// TIA Portal project "261019_Kommissionierung_GA_Analog2_20261019_1400" (V17)

(* hardware
DEVICE "S7300/ET200M-Station_1"  S7-300 station
   slot 0: "Profilschiene_0"  Rail  6ES7 390-1***0-0AA0
   slot 1: "PS 307 5A_1"  PS 307 5A  6ES7 307-1EA01-0AA0
   slot 2: "PLC_WBS_Bus_1"  CPU 314C-2 DP  6ES7 314-6CH04-0AB0  V3.3
      slot 0: "MPI-Schnittstelle_1"  MPI
      slot 1: "DP-Schnittstelle_1"  DP
      slot 2: "DI 24/DO 16_1"  DI24/DO16
      slot 3: "AI 5/AO 2_1"  AI5/AO2
      slot 4: "Zählen_1"  Counter
      slot 5: "Positionieren_1"  Positioning
   slot 4: "DI 64x24VDC sinking/souring_1"  DI64 x 24VDC  6ES7 321-1BP00-0AA0
   slot 5: "DI 64x24VDC sinking/souring_2"  DI64 x 24VDC  6ES7 321-1BP00-0AA0
   slot 6: "DI 64x24VDC sinking/souring_3"  DI64 x 24VDC  6ES7 321-1BP00-0AA0
   slot 7: "DI 64x24VDC sinking/souring_4"  DI64 x 24VDC  6ES7 321-1BP00-0AA0
   slot 8: "DO 64x24VDC/0.3A sourcing_1"  DO64 x 24VDC / 0.3A, P  6ES7 322-1BP00-0AA0
   slot 9: "DO 64x24VDC/0.3A sourcing_2"  DO64 x 24VDC / 0.3A, P  6ES7 322-1BP00-0AA0
   slot 10: "DO 64x24VDC/0.3A sourcing_3"  DO64 x 24VDC / 0.3A, P  6ES7 322-1BP00-0AA0
   slot 11: "DO 64x24VDC/0.3A sourcing_4"  DO64 x 24VDC / 0.3A, P  6ES7 322-1BP00-0AA0
*)

// ===== PLC "PLC_WBS_Bus_1"  CPU 314C-2 DP =====

VAR_GLOBAL   // PLC tag table "Standard-Variablentabelle"
   "NotAusOK" AT %M20.0 : Bool;
   "Band 1 Grün" AT %M41.0 : Bool;
   "Band 2 Blau" AT %M40.1 : Bool;
   "Signal_Start_Bearbeitung" AT %M80.0 : Bool;
   "Band 3 Blau" AT %M40.3 : Bool;
   "Auswahl Unterteil Blau" AT %M42.0 : Bool;
   "Band 6 Blau" AT %M40.4 : Bool;
   "Klemmen UT" AT %M80.2 : Bool;
   "Klemmen Unterteil Blau" AT %M44.0 : Bool;
   "Auswahl Oberteil Blau" AT %M42.1 : Bool;
   "Klemmen Oberteil Blau" AT %M44.1 : Bool;
   "Klemmen OT" AT %M80.3 : Bool;
   "Freigabe_Zusammenbau UT Blau" AT %M82.0 : Bool;
   "Freigabe_Zusammenbau OT Blau" AT %M82.1 : Bool;
   "Teil in Pos. nf" AT %M81.0 : Bool;
   "Teil in Pos. pf" AT %M81.1 : Bool;
   "Z-Achse Greifer Blau" AT %M82.2 : Bool;
   "Greifer Blau" AT %M82.3 : Bool;
   "X-Achse Greifer" AT %M82.4 : Bool;
   "Sensor Weitergabe pf Blau" AT %M82.6 : Bool;
   "Sensor Weitergabe pf 2 Blau" AT %M82.7 : Bool;
   "Start Zusammenbau Blau" AT %M83.0 : Bool;
   "Start zusammen bau pf Blau" AT %M83.3 : Bool;
   "Greifer X-Achse Blau" AT %M83.4 : Bool;
   "Z-Achse senken Zusammenbau" AT %M83.5 : Bool;
   "Teil erkannt pf Blau" AT %M83.7 : Bool;
   "Zusammenbau fertig" AT %M84.6 : Bool;
   "FreigabeKommissionierung Blau" AT %M90.0 : Bool;
   "Anlage Freigegeben" AT %M1.0 : Bool;
   "2Hz" AT %M100.3 : Bool;
   "Betriebsbereit" AT %M20.1 : Bool;
   "Anlage An" AT %M20.2 : Bool;
   "Warnung" AT %M20.3 : Bool;
   "T10s" AT %M20.4 : Bool;
   "Betriebsbereit pf" AT %M20.5 : Bool;
   "Objekt erzeugen Blau" AT %M20.6 : Bool;
   "Start Allgemein" AT %M20.7 : Bool;
   "Start pf" AT %M21.0 : Bool;
   "Auswahl OT_UT Blau" AT %M92.0 : Bool;
   "Start_Signal" AT %M21.2 : Bool;
   "Greifer nf Blau" AT %M83.2 : Bool;
   "X-Achse pf" AT %M84.3 : Bool;
   "Teil erkannt pf(1)" AT %M79.0 : Bool;
   "Start Zusammenbau pf" AT %M81.2 : Bool;
   "Teil fertig Blau" AT %M84.4 : Bool;
   "Grundstellung Roboter Blau" AT %M84.7 : Bool;
   "Teil fertig SR Blau" AT %M85.0 : Bool;
   "Emmit pf" AT %M21.4 : Bool;
   "TB3006 pf" AT %M40.2 : Bool;
   "Start  t1s. pf Blau" AT %M19.1 : Bool;
   "Neues Objekt pf Blau" AT %M19.2 : Bool;
   "Signal_Start_Bearbeitung Grün" AT %M80.1 : Bool;
   "Band 2 Grün" AT %M40.0 : Bool;
   "TB 4006 pf" AT %M40.5 : Bool;
   "Band 3 Grün" AT %M40.6 : Bool;
   "Auswahl Oberteil Grün" AT %M40.7 : Bool;
   "Auswahl Unterteil Grün" AT %M41.1 : Bool;
   "Teil vor Pos. nf" AT %M81.4 : Bool;
   "Klemmen Oberteil Grün" AT %M44.2 : Bool;
   "Teil in Pos. nf Grün" AT %M81.3 : Bool;
   "Klemmen Unterteil Grün" AT %M44.3 : Bool;
   "Band 6 Grün" AT %M41.2 : Bool;
   "FreigabeKommissionierung Grün" AT %M90.1 : Bool;
   "Freigabe_Zusammenbau UT Grün" AT %M84.0 : Bool;
   "Sensor Weitergabe pf Grün" AT %M80.4 : Bool;
   "Freigabe_Zusammenbau OT Grün" AT %M84.1 : Bool;
   "Sensor Weitergabe pf 2 Grün" AT %M84.5 : Bool;
   "Start Zusammenbau Grün" AT %M83.1 : Bool;
   "Start zusammen bau pf Grün" AT %M83.6 : Bool;
   "X-Achse pf Grün" AT %M85.1 : Bool;
   "Z-Achse Greifer Grün" AT %M85.2 : Bool;
   "Greifer X-Achse Grün" AT %M85.3 : Bool;
   "Teil erkannt pf Grün" AT %M85.4 : Bool;
   "Teil erkannt pf(1) Grün" AT %M85.5 : Bool;
   "Teil fertig Grün" AT %M85.6 : Bool;
   "Greifer Grün" AT %M85.7 : Bool;
   "Start Zusammenbau pf Grün" AT %M90.2 : Bool;
   "Greifer nf Grün" AT %M90.3 : Bool;
   "Greifer X-Achse Grün(1)" AT %M90.4 : Bool;
   "Teil erkannt pf Grün(1)" AT %M90.5 : Bool;
   "Teil fertig SR Grün" AT %M90.6 : Bool;
   "Grundstellung Roboter Grün" AT %M90.7 : Bool;
   "FreigabeKommissionierung Grün(1)" AT %M92.1 : Bool;
   "Auswahl OT_UT Grün" AT %M92.2 : Bool;
   "Start  t1s. pf Grün" AT %M19.3 : Bool;
   "Neues Objekt pf Grün" AT %M19.4 : Bool;
   "Objekt erzeugen Grün" AT %M19.5 : Bool;
END_VAR

VAR_GLOBAL   // PLC tag table "Betriebsart"
   "S0_HS" AT %E0.0 : Bool;   // Hauptschalter 0-Aus, 1-Ein
   "S1_Not_Halt" AT %E0.1 : Bool;   // Not-Halt NC
   "S2_START" AT %E0.2 : Bool;   // Taster START NO
   "S3_STOP" AT %E0.3 : Bool;   // Taster STOP NC
   "Res_E04" AT %E0.4 : Bool;
   "Res_E05" AT %E0.5 : Bool;
   "Res_E06" AT %E0.6 : Bool;
   "Res_E07" AT %E0.7 : Bool;
   "Res_E10" AT %E1.0 : Bool;
   "Res_E11" AT %E1.1 : Bool;
   "Res_E12" AT %E1.2 : Bool;
   "Res_E13" AT %E1.3 : Bool;
   "Res_E14" AT %E1.4 : Bool;
   "Res_E15" AT %E1.5 : Bool;
   "Res_E16" AT %E1.6 : Bool;
   "Factory_IO_RUN" AT %E1.7 : Bool;   // Rückmeldung Factory IO läuft
   "P1_MS_RT" AT %A0.0 : Bool;   // Meldesäule Rot
   "P2_MS_GE" AT %A0.1 : Bool;   // Meldesäule Gelb
   "P3_MS_GN" AT %A0.2 : Bool;   // Meldesäule Grün
   "P10_START" AT %A0.3 : Bool;   // Anzeige grün in START-Taster
   "P11_STOP" AT %A0.4 : Bool;   // Anzeige gelb in START-Taster
   "Res_A0.5" AT %A0.5 : Bool;
   "P12_Anfahrwarnung" AT %A0.6 : Bool;   // Rundumleuchte System
   "P13_Sirene" AT %A0.7 : Bool;   // Sirene System
   "Res_A10" AT %A1.0 : Bool;
   "Res_A11" AT %A1.1 : Bool;
   "Res_A12" AT %A1.2 : Bool;
   "Res_A13" AT %A1.3 : Bool;
   "Res_A14" AT %A1.4 : Bool;
   "Res_A15" AT %A1.5 : Bool;
   "Res_A16" AT %A1.6 : Bool;
   "Res_A17" AT %A1.7 : Bool;
   "Log_1" AT %M0.1 : Bool;   // statisch "1"
   "Log_0" AT %M0.0 : Bool;   // statisch "0"
   "Takt_1HZ" AT %M100.5 : Bool;   // Taktmerker 1 Hz
   "Anzeige_Anzahl_Teile_BL" AT %AW22 : Int;   // Anzeige Teile blau im Lager
   "Anzeige_Anzahl_Teile_GN" AT %AW24 : Int;   // Anzeige Teile grün im Lager
   "Reset Nothalt" AT %M0.2 : Bool;
END_VAR

VAR_GLOBAL   // PLC tag table "Montage"
   "B3001_TB3001" AT %E2.0 : Bool;   // Transportband-Ende NC
   "B3002_TB3001" AT %E2.1 : Bool;   // Teil nachPositionierer NC
   "B3003_Teil_vor_POS" AT %E2.2 : Bool;   // Teil vor Positionierer NC
   "B3004_TB3001" AT %E2.3 : Bool;   // Transportband-Anfang NC
   "B3005_TB3002" AT %E2.4 : Bool;   // Transportband-Ende NC
   "B3006_TB3006" AT %E2.5 : Bool;   // Teil vor Schwenkarm NC
   "B3007_UT_BL" AT %E2.6 : Bool;   // Farbsensor Erkennung Farbteil Unterteil blau
   "B3008_OT_BL" AT %E2.7 : Bool;   // Farbsensor Erkennung Farbteil Oberteil blau
   "B3009_TB3006" AT %E3.0 : Bool;   // Transportband-Anfang NC
   "B3010_TB3007" AT %E3.1 : Bool;   // Transportband-Ende NC
   "B3011_TB3007" AT %E3.2 : Bool;   // Transportband-Anfang NC
   "B3012_TB3008" AT %E3.3 : Bool;   // Transportband-Ende NC
   "B3013_TB3008" AT %E3.4 : Bool;   // Transportband-Anfang NC
   "B3014_TB3005" AT %E3.5 : Bool;   // Transportband-Anfang NC
   "B3015_TB3005" AT %E3.6 : Bool;   // Transportband-Ende
   "B3016_TB3004" AT %E3.7 : Bool;   // Transportband-Anfang
   "B3017_Teil_vor_POS" AT %E4.0 : Bool;   // Teil vor Positionierer NC
   "B3018_TB3004" AT %E4.1 : Bool;   // Transportband-Ende NC
   "B3030_POS3001_geklemmt" AT %E4.2 : Bool;   // Positionierer RM geklemmt
   "B3031_POS3001_Heben_Senken" AT %E4.3 : Bool;   // Positionierer RM Bewegung
   "B3040_POS3002_geklemmt" AT %E4.4 : Bool;   // Positionierer RM geklemmt
   "B3041_POS3002_Heben_Senken" AT %E4.5 : Bool;   // Positionierer RM Bewegung
   "Res_E46" AT %E4.6 : Bool;
   "Res_E47" AT %E4.7 : Bool;
   "B3050_PAP3001_RM_X" AT %E5.0 : Bool;
   "B3051_PAP3001_RM_Z" AT %E5.1 : Bool;
   "B3052_PAP3001_Teil_erkannt" AT %E5.2 : Bool;
   "B3070_FZ_3001_Busy" AT %E5.3 : Bool;
   "B3071_FZ_3001_Error" AT %E5.4 : Bool;
   "B3072_FZ_Tür_offen" AT %E5.5 : Bool;
   "Res_E56" AT %E5.6 : Bool;
   "Res_E57" AT %E5.7 : Bool;
   "B4001_TB4001" AT %E6.0 : Bool;   // Transportband-Ende NC
   "B4002_TB4001" AT %E6.1 : Bool;   // Teil nachPositionierer NC
   "B4003_Teil_vor_POS" AT %E6.2 : Bool;   // Teil vor Positionierer NC
   "B4004_TB4001" AT %E6.3 : Bool;   // Transportband-Anfang NC
   "B4005_TB4002" AT %E6.4 : Bool;   // Transportband-Ende NC
   "B4006_TB4006" AT %E6.5 : Bool;   // Teil vor Schwenkarm NC
   "B4007_UT_GN" AT %E6.6 : Bool;   // Farbsensor Erkennung Farbteil Unterteil blau
   "B4008_OT_GN" AT %E6.7 : Bool;   // Farbsensor Erkennung Farbteil Oberteil blau
   "B4009_TB4006" AT %E7.0 : Bool;   // Transportband-Anfang NC
   "B4010_TB4007" AT %E7.1 : Bool;   // Transportband-Ende NC
   "B4011_TB4007" AT %E7.2 : Bool;   // Transportband-Anfang NC
   "B4012_TB4008" AT %E7.3 : Bool;   // Transportband-Ende NC
   "B4013_TB4008" AT %E7.4 : Bool;   // Transportband-Anfang NC
   "B4014_TB4005" AT %E7.5 : Bool;   // Transportband-Anfang NC
   "B4015_TB4005" AT %E7.6 : Bool;   // Transportband-Ende
   "B4016_TB4004" AT %E7.7 : Bool;   // Transportband-Anfang
   "B4017_Teil_vor_POS" AT %E8.0 : Bool;   // Teil vor Positionierer NC
   "B4018_TB4004" AT %E8.1 : Bool;   // Transportband-Ende NC
   "B4030_POS4001_geklemmt" AT %E8.2 : Bool;   // Positionierer RM geklemmt
   "B4031_POS4001_Heben_Senken" AT %E8.3 : Bool;   // Positionierer RM Bewegung
   "B4040_POS4002_geklemmt" AT %E8.4 : Bool;   // Positionierer RM geklemmt
   "B4041_POS4002_Heben_Senken" AT %E8.5 : Bool;   // Positionierer RM Bewegung
   "Res_E86" AT %E8.6 : Bool;
   "Res_E87" AT %E8.7 : Bool;
   "B4050_PAP4001_RM_X" AT %E9.0 : Bool;   // Pick-and-Place X-aktiv
   "B4051_PAP4001_RM_Z" AT %E9.1 : Bool;   // Pick-and-Place Z-aktiv
   "B4052_PAP4001_Teil_erkannt" AT %E9.2 : Bool;   // Teil am Greifer erkannt
   "B4070_FZ_4001_Busy" AT %E9.3 : Bool;   // Fertigungszentrum
   "B4071_FZ_4001_Error" AT %E9.4 : Bool;   // Fertigungszentrum
   "B4072_FZ_4001_Tür_offen" AT %E9.5 : Bool;   // Fertigungszentrum
   "Res_E96" AT %E9.6 : Bool;
   "Res_E97" AT %E9.7 : Bool;
   "TB3001" AT %A2.0 : Bool;
   "TB3002" AT %A2.1 : Bool;
   "TB3003" AT %A2.2 : Bool;
   "TB3004" AT %A2.3 : Bool;
   "TB3005" AT %A2.4 : Bool;
   "TB3006" AT %A2.5 : Bool;
   "TB3007" AT %A2.6 : Bool;
   "TB3008" AT %A2.7 : Bool;
   "FZ_3001_Start" AT %A3.0 : Bool;   // Fertigungszentrum Start
   "FZ_3001_Stop" AT %A3.1 : Bool;   // Fertigungszentrum Stop
   "FZ_3001_OT_UT" AT %A3.2 : Bool;   // Fertigungszentrum UT =0 / OT=1
   "Sorter_Arm_3001_schwenken" AT %A3.3 : Bool;
   "Sorter_Arm_3001_Band_V" AT %A3.4 : Bool;
   "Sorter_Arm_3001_Band_R" AT %A3.5 : Bool;
   "POS3001_Klemmen" AT %A3.6 : Bool;
   "POS3001_Heben" AT %A3.7 : Bool;
   "POS3002_Klemmen" AT %A4.0 : Bool;
   "POS3002_Heben" AT %A4.1 : Bool;
   "PAP3001_X" AT %A4.2 : Bool;
   "PAP3001_Z" AT %A4.3 : Bool;
   "PAP3001_Greifer" AT %A4.4 : Bool;
   "STOP_3001" AT %A4.5 : Bool;
   "Res_A46" AT %A4.6 : Bool;
   "Emitter_1 Blau" AT %A4.7 : Bool;   // Emitter_1
   "TB4001" AT %A5.0 : Bool;
   "TB4002" AT %A5.1 : Bool;
   "TB4003" AT %A5.2 : Bool;
   "TB4004" AT %A5.3 : Bool;
   "TB4005" AT %A5.4 : Bool;
   "TB4006" AT %A5.5 : Bool;
   "TB4007" AT %A5.6 : Bool;
   "TB4008" AT %A5.7 : Bool;
   "FZ_4001_Start" AT %A6.0 : Bool;   // Fertigungszentrum Start
   "FZ_4001_Stop" AT %A6.1 : Bool;   // Fertigungszentrum Stop
   "FZ_4001_OT_UT" AT %A6.2 : Bool;   // Fertigungszentrum UT =0 / OT=1
   "Sorter_Arm_4001_schwenken" AT %A6.3 : Bool;
   "Sorter_Arm_4001_Band_V" AT %A6.4 : Bool;
   "Sorter_Arm_4001_Band_R" AT %A6.5 : Bool;
   "POS4001_Klemmen" AT %A6.6 : Bool;
   "POS4001_Heben" AT %A6.7 : Bool;
   "POS4002_Klemmen" AT %A7.0 : Bool;
   "POS4002_Heben" AT %A7.1 : Bool;
   "PAP4001_X" AT %A7.2 : Bool;
   "PAP4001_Z" AT %A7.3 : Bool;
   "PAP4001_Greifer" AT %A7.4 : Bool;
   "STOP4001" AT %A7.5 : Bool;
   "Res_A76" AT %A7.6 : Bool;
   "Emitter_2 Grün" AT %A7.7 : Bool;
   "FZ_3001_Bearbeitungszeit" AT %EW20 : Int;
   "FZ_4001_Bearbeitungszeit" AT %EW22 : Int;
END_VAR

VAR_GLOBAL   // PLC tag table "Kommisionierung"
   "B5001_TB5001" AT %E10.0 : Bool;   // Teil vom Emitter vorhanden
   "B5002_TB5001" AT %E10.1 : Bool;   // Transportband-Ende
   "B5003_TB5002" AT %E10.2 : Bool;   // Transportband-Anfang
   "B5004_TB5002" AT %E10.3 : Bool;   // Transportband-Ende
   "B5005_TB5003" AT %E10.4 : Bool;   // Transportband-Anfang
   "B5006_TB5003" AT %E10.5 : Bool;   // Transportband-Ende
   "B5007_TB5004" AT %E10.6 : Bool;   // Transportband-Anfang
   "B5008_TB5004" AT %E10.7 : Bool;   // Transportband-Ende
   "B5009_TB5005" AT %E11.0 : Bool;   // Transportband-Anfang
   "B5010_TB5005" AT %E11.1 : Bool;   // Transportband-Ende
   "B5011_Farbteil_GN" AT %E11.2 : Bool;   // Farberkennung GN
   "B5012_Farbteil_BL" AT %E11.3 : Bool;   // Farberkennung_BL
   "B5013_TB5006" AT %E11.4 : Bool;   // Transportband-Anfang
   "B5014_TB5006" AT %E11.5 : Bool;   // Transportband-Ende blaue Produkte
   "B5016_Teil_vorhanden" AT %E11.7 : Bool;   // Teil vom Emitter generiert
   "B5018_Teil_vorhanden" AT %E12.1 : Bool;   // Teil vom Emitter generiert
   "B5019_TB5009" AT %E12.2 : Bool;   // Transportband-Anfang
   "B5020_TB5009" AT %E12.3 : Bool;   // Transportband-Ende
   "B5021_TB5010" AT %E12.4 : Bool;   // Transportband-Anfang
   "B5022_TB5010" AT %E12.5 : Bool;   // Transportband-Ende grüne Produkte
   "Res_E126" AT %E12.6 : Bool;
   "Res_E127" AT %E12.7 : Bool;
   "B5030_PAP5001_RM_X" AT %E13.0 : Bool;
   "B5031_PAP5001_RM_Z" AT %E13.1 : Bool;
   "B5032_PAP5001_Teil_erkannt" AT %E13.2 : Bool;
   "B5040_PAP5002_RM_X" AT %E13.3 : Bool;
   "B5041_PAP5002_RM_Z" AT %E13.4 : Bool;
   "B5042_PAP5002_Teil_erkannt" AT %E13.5 : Bool;
   "Res_E136" AT %E13.6 : Bool;
   "Res_E137" AT %E13.7 : Bool;
   "TB5001" AT %A8.0 : Bool;
   "TB5002" AT %A8.1 : Bool;
   "TB5003" AT %A8.2 : Bool;
   "TB5004" AT %A8.3 : Bool;
   "TB5005" AT %A8.4 : Bool;
   "TB5006" AT %A8.5 : Bool;
   "TB5007" AT %A8.6 : Bool;
   "TB5008" AT %A8.7 : Bool;
   "TB5009" AT %A9.0 : Bool;
   "TB5010" AT %A9.1 : Bool;
   "STOP5001" AT %A9.2 : Bool;   // Stopper
   "STOP5002" AT %A9.3 : Bool;   // Stopper
   "STOP5003" AT %A9.4 : Bool;   // Stopper
   "STOP5004" AT %A9.5 : Bool;   // Stopper
   "STOP5005" AT %A9.6 : Bool;   // Stopper
   "Res_A97" AT %A9.7 : Bool;
   "PAP5001_X" AT %A10.0 : Bool;
   "PAP5001_Z" AT %A10.1 : Bool;
   "PAP5001_Greifer" AT %A10.2 : Bool;
   "PAP5002_X" AT %A10.3 : Bool;
   "PAP5002_Z" AT %A10.4 : Bool;
   "PAP5002_Greifer" AT %A10.5 : Bool;
   "Res_A106" AT %A10.6 : Bool;
   "Res_A107" AT %A10.7 : Bool;
   "RS5001_V" AT %A11.0 : Bool;   // Rollensorter Antrieb ein
   "RS5001_links" AT %A11.1 : Bool;   // Rollensorter Steuerung links
   "RS5001_rechts" AT %A11.2 : Bool;   // Rollensorter Steuerung rechts
   "Res_A113" AT %A11.3 : Bool;
   "Res_A114" AT %A11.4 : Bool;
   "Emitter_1" AT %A11.5 : Bool;
   "Emitter_2" AT %A11.6 : Bool;
   "Emitter_3" AT %A11.7 : Bool;
   "TA_P&P2_SetPoint_X" AT %AW24 : Int;
   "TA_P&P2_SetPoint_Z" AT %AW26 : Int;
   "TA_P&P1_SetPoint_X" AT %AW20 : Int;
   "TA_P&P1_SetPoint_Z" AT %AW22 : Int;
   "TA_P&P2_Pos_X" AT %EW24 : Int;
   "TA_P&P2_Pos_Z" AT %EW26 : Int;
   "TA_P&P1_Pos_X" AT %EW20 : Int;
   "TA_P&P1_Pos_Z" AT %EW22 : Int;
   "B5015_Teil_in_Pos" AT %E11.6 : Bool;
   "B5017_Teil_in_Pos" AT %E12.0 : Bool;
END_VAR

// folder: Kommissionierung

DATA_BLOCK "100_DB_Kommissionierung"   // DB100
{ S7_Optimized_Access := 'FALSE' }
VERSION : 0.1
   VAR
      xNotAusOK : Bool;
      xAnlageAusgeschaltet : Bool;
      xAnlageStartet : Bool;
      xAnlageEin : Bool;
      xGA1_Fertig : Bool;
      xGA2_Fertig : Bool;
      strGA1_Meldung : String[30];
      strGA2_Meldung : String[30];
      iIndex_Förderband : Int;
   END_VAR
BEGIN
END_DATA_BLOCK

// folder: Kommissionierung/iDB

DATA_BLOCK "02_AnlageEinAus_DB"   // DB29
{ S7_Optimized_Access := 'FALSE' }
VERSION : 0.1
// stored: InstanceOfName 02_AnlageEinAus
"02_AnlageEinAus"
BEGIN
END_DATA_BLOCK

DATA_BLOCK "03_Förderband_DB"   // DB30
{ S7_Optimized_Access := 'FALSE' }
VERSION : 0.1
// stored: InstanceOfName 03_Förderband
"03_Förderband"
BEGIN
END_DATA_BLOCK

DATA_BLOCK "04_Greifarm_DB"   // DB31
{ S7_Optimized_Access := 'FALSE' }
VERSION : 0.1
// stored: InstanceOfName 04_Greifarm
"04_Greifarm"
BEGIN
END_DATA_BLOCK

DATA_BLOCK "04_Greifarm_DB_1"   // DB32
{ S7_Optimized_Access := 'FALSE' }
VERSION : 0.1
// stored: InstanceOfName 04_Greifarm
"04_Greifarm"
BEGIN
END_DATA_BLOCK

// folder: Montage/Bearbeitung Blau

DATA_BLOCK "01_Transportband vor Bearbeitung_DB"   // DB1
{ S7_Optimized_Access := 'FALSE' }
VERSION : 0.1
// stored: InstanceOfName 01Transportband vor Bearbeitung
"01Transportband vor Bearbeitung"
BEGIN
END_DATA_BLOCK

DATA_BLOCK "Bearbeitung_DB"   // DB2
{ S7_Optimized_Access := 'FALSE' }
VERSION : 0.1
// stored: InstanceOfName 02_Bearbeitung
"02_Bearbeitung"
BEGIN
END_DATA_BLOCK

DATA_BLOCK "02_Bearbeitung_DB"   // DB3
{ S7_Optimized_Access := 'FALSE' }
VERSION : 0.1
// stored: InstanceOfName 02_Bearbeitung
"02_Bearbeitung"
BEGIN
END_DATA_BLOCK

DATA_BLOCK "03_Weiterverarbeitung_DB"   // DB4
{ S7_Optimized_Access := 'FALSE' }
VERSION : 0.1
// stored: InstanceOfName 03_Weiterverarbeitung
"03_Weiterverarbeitung"
BEGIN
END_DATA_BLOCK

DATA_BLOCK "04_Zusammenbau_DB"   // DB6
{ S7_Optimized_Access := 'FALSE' }
VERSION : 0.1
// stored: InstanceOfName 04_Zusammenbau
"04_Zusammenbau"
BEGIN
END_DATA_BLOCK

DATA_BLOCK "05_Weitergabe_DB"   // DB11
{ S7_Optimized_Access := 'FALSE' }
VERSION : 0.1
// stored: InstanceOfName 05_Weitergabe
"05_Weitergabe"
BEGIN
END_DATA_BLOCK

DATA_BLOCK "06_Auswahl OT_UT_DB"   // DB15
{ S7_Optimized_Access := 'FALSE' }
VERSION : 0.1
// stored: InstanceOfName 06_Auswahl OT_UT
"06_Auswahl OT_UT"
BEGIN
END_DATA_BLOCK

// folder: Montage/Bearbeitung Grün

DATA_BLOCK "01_Transportband vor Bearbeitung_DB_Grün"   // DB20
{ S7_Optimized_Access := 'FALSE' }
VERSION : 0.1
// stored: InstanceOfName 01Transportband vor Bearbeitung Grün
"01Transportband vor Bearbeitung Grün"
BEGIN
END_DATA_BLOCK

DATA_BLOCK "Bearbeitung_DB_Grün"   // DB21
{ S7_Optimized_Access := 'FALSE' }
VERSION : 0.1
// stored: InstanceOfName 02_Bearbeitung Grün
"02_Bearbeitung Grün"
BEGIN
END_DATA_BLOCK

DATA_BLOCK "02_Bearbeitung_DB_Grün"   // DB22
{ S7_Optimized_Access := 'FALSE' }
VERSION : 0.1
// stored: InstanceOfName 02_Bearbeitung Grün
"02_Bearbeitung Grün"
BEGIN
END_DATA_BLOCK

DATA_BLOCK "03_Weiterverarbeitung_DB_Grün"   // DB23
{ S7_Optimized_Access := 'FALSE' }
VERSION : 0.1
// stored: InstanceOfName 03_Weiterverarbeitung Grün
"03_Weiterverarbeitung Grün"
BEGIN
END_DATA_BLOCK

DATA_BLOCK "04_Zusammenbau_DB_Grün"   // DB24
{ S7_Optimized_Access := 'FALSE' }
VERSION : 0.1
// stored: InstanceOfName 04_Zusammenbau Grün
"04_Zusammenbau Grün"
BEGIN
END_DATA_BLOCK

DATA_BLOCK "05_Weitergabe_DB_Grün"   // DB25
{ S7_Optimized_Access := 'FALSE' }
VERSION : 0.1
// stored: InstanceOfName 05_Weitergabe Grün
"05_Weitergabe Grün"
BEGIN
END_DATA_BLOCK

DATA_BLOCK "06_Auswahl OT_UT_DB_Grün"   // DB26
{ S7_Optimized_Access := 'FALSE' }
VERSION : 0.1
// stored: InstanceOfName 06_Auswahl OT_UT_Grün
"06_Auswahl OT_UT_Grün"
BEGIN
END_DATA_BLOCK

// folder: Montage/iDB

DATA_BLOCK "05_Weitergabe_DB_1"   // DB5
{ S7_Optimized_Access := 'FALSE' }
VERSION : 0.1
// stored: InstanceOfName 05_Weitergabe
"05_Weitergabe"
BEGIN
END_DATA_BLOCK

DATA_BLOCK "01Transportband vor Bearbeitung Grün_DB"   // DB9
{ S7_Optimized_Access := 'FALSE' }
VERSION : 0.1
// stored: InstanceOfName 01Transportband vor Bearbeitung Grün
"01Transportband vor Bearbeitung Grün"
BEGIN
END_DATA_BLOCK

DATA_BLOCK "02_Bearbeitung Grün_DB"   // DB10
{ S7_Optimized_Access := 'FALSE' }
VERSION : 0.1
// stored: InstanceOfName 02_Bearbeitung Grün
"02_Bearbeitung Grün"
BEGIN
END_DATA_BLOCK

DATA_BLOCK "03_Weiterverarbeitung Grün_DB"   // DB14
{ S7_Optimized_Access := 'FALSE' }
VERSION : 0.1
// stored: InstanceOfName 03_Weiterverarbeitung Grün
"03_Weiterverarbeitung Grün"
BEGIN
END_DATA_BLOCK

DATA_BLOCK "04_Zusammenbau Grün_DB"   // DB16
{ S7_Optimized_Access := 'FALSE' }
VERSION : 0.1
// stored: InstanceOfName 04_Zusammenbau Grün
"04_Zusammenbau Grün"
BEGIN
END_DATA_BLOCK

DATA_BLOCK "05_Weitergabe Grün_DB"   // DB17
{ S7_Optimized_Access := 'FALSE' }
VERSION : 0.1
// stored: InstanceOfName 05_Weitergabe Grün
"05_Weitergabe Grün"
BEGIN
END_DATA_BLOCK

DATA_BLOCK "06_Auswahl OT_UT_Grün_DB"   // DB18
{ S7_Optimized_Access := 'FALSE' }
VERSION : 0.1
// stored: InstanceOfName 06_Auswahl OT_UT_Grün
"06_Auswahl OT_UT_Grün"
BEGIN
END_DATA_BLOCK

DATA_BLOCK "00_Startbedingungen_2_DB"   // DB27
{ S7_Optimized_Access := 'FALSE' }
VERSION : 0.1
// stored: InstanceOfName 00_Startbedingungen_2
"00_Startbedingungen_2"
BEGIN
END_DATA_BLOCK

// folder: (top level)

ORGANIZATION_BLOCK "Main"   // OB1, FBD
TITLE = "Main Program Sweep (Cycle)"
{ S7_Optimized_Access := 'FALSE' }
VERSION : 0.1
   VAR_TEMP
      OB1_EV_CLASS : Byte;   // Bits 0-3 = 1 (Coming event), Bits 4-7 = 1 (Event class 1)
      OB1_SCAN_1 : Byte;   // 1 (Cold restart scan 1 of OB 1), 3 (Scan 2-n of OB 1)
      OB1_PRIORITY : Byte;   // Priority of OB Execution
      OB1_OB_NUMBR : Byte;   // 1 (Organization block 1, OB1)
      OB1_RESERVED_1 : Byte;   // Reserved for system
      OB1_RESERVED_2 : Byte;   // Reserved for system
      OB1_PREV_CYCLE : Int;   // Cycle time of previous OB1 scan (milliseconds)
      OB1_MIN_CYCLE : Int;   // Minimum cycle time of OB1 (milliseconds)
      OB1_MAX_CYCLE : Int;   // Maximum cycle time of OB1 (milliseconds)
      OB1_DATE_TIME : Date_And_Time;   // Date and time OB1 started
   END_VAR
BEGIN

REGION Network 1: Startbedingung
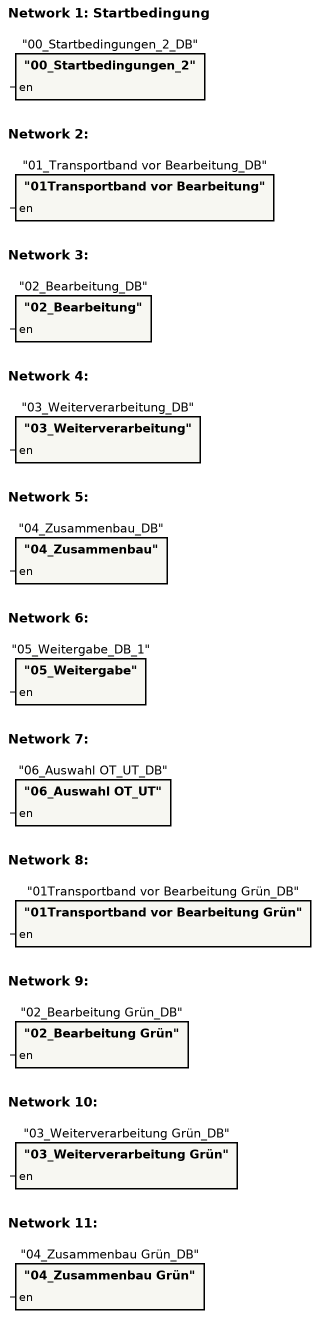
   "00_Startbedingungen_2_DB"();   // "00_Startbedingungen_2"
END_REGION

REGION Network 2
   "01_Transportband vor Bearbeitung_DB"();   // "01Transportband vor Bearbeitung"
END_REGION

REGION Network 3
   "02_Bearbeitung_DB"();   // "02_Bearbeitung"
END_REGION

REGION Network 4
   "03_Weiterverarbeitung_DB"();   // "03_Weiterverarbeitung"
END_REGION

REGION Network 5
   "04_Zusammenbau_DB"();   // "04_Zusammenbau"
END_REGION

REGION Network 6
   "05_Weitergabe_DB_1"();   // "05_Weitergabe"
END_REGION

REGION Network 7
   "06_Auswahl OT_UT_DB"();   // "06_Auswahl OT_UT"
END_REGION

REGION Network 8
   "01Transportband vor Bearbeitung Grün_DB"();   // "01Transportband vor Bearbeitung Grün"
END_REGION

REGION Network 9
   "02_Bearbeitung Grün_DB"();   // "02_Bearbeitung Grün"
END_REGION

REGION Network 10
   "03_Weiterverarbeitung Grün_DB"();   // "03_Weiterverarbeitung Grün"
END_REGION

REGION Network 11
   "04_Zusammenbau Grün_DB"();   // "04_Zusammenbau Grün"
END_REGION

REGION Network 12
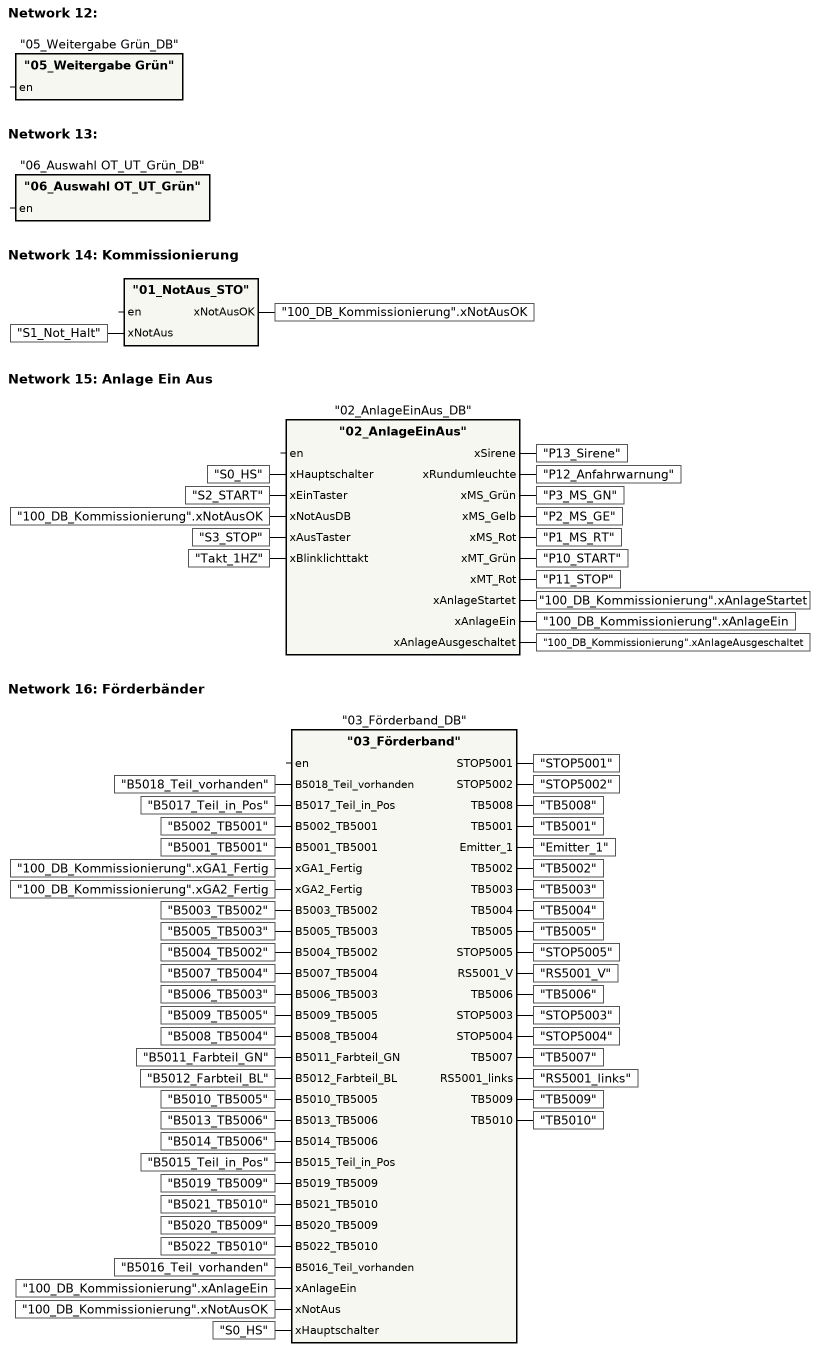
   "05_Weitergabe Grün_DB"();   // "05_Weitergabe Grün"
END_REGION

REGION Network 13
   "06_Auswahl OT_UT_Grün_DB"();   // "06_Auswahl OT_UT_Grün"
END_REGION

REGION Network 14: Kommissionierung
   "01_NotAus_STO"(xNotAus := "S1_Not_Halt", xNotAusOK => "100_DB_Kommissionierung".xNotAusOK);
END_REGION

REGION Network 15: Anlage Ein Aus
   "02_AnlageEinAus_DB"(xHauptschalter := "S0_HS",   // "02_AnlageEinAus"
                        xEinTaster := "S2_START",
                        xNotAusDB := "100_DB_Kommissionierung".xNotAusOK,
                        xAusTaster := "S3_STOP",
                        xBlinklichttakt := "Takt_1HZ",
                        xSirene => "P13_Sirene",
                        xRundumleuchte => "P12_Anfahrwarnung",
                        xMS_Grün => "P3_MS_GN",
                        xMS_Gelb => "P2_MS_GE",
                        xMS_Rot => "P1_MS_RT",
                        xMT_Grün => "P10_START",
                        xMT_Rot => "P11_STOP",
                        xAnlageStartet => "100_DB_Kommissionierung".xAnlageStartet,
                        xAnlageEin => "100_DB_Kommissionierung".xAnlageEin,
                        xAnlageAusgeschaltet => "100_DB_Kommissionierung".xAnlageAusgeschaltet);
END_REGION

REGION Network 16: Förderbänder
   "03_Förderband_DB"(B5018_Teil_vorhanden := "B5018_Teil_vorhanden",   // "03_Förderband"
                      B5017_Teil_in_Pos := "B5017_Teil_in_Pos",
                      B5002_TB5001 := "B5002_TB5001",
                      B5001_TB5001 := "B5001_TB5001",
                      xGA1_Fertig := "100_DB_Kommissionierung".xGA1_Fertig,
                      xGA2_Fertig := "100_DB_Kommissionierung".xGA2_Fertig,
                      B5003_TB5002 := "B5003_TB5002",
                      B5005_TB5003 := "B5005_TB5003",
                      B5004_TB5002 := "B5004_TB5002",
                      B5007_TB5004 := "B5007_TB5004",
                      B5006_TB5003 := "B5006_TB5003",
                      B5009_TB5005 := "B5009_TB5005",
                      B5008_TB5004 := "B5008_TB5004",
                      B5011_Farbteil_GN := "B5011_Farbteil_GN",
                      B5012_Farbteil_BL := "B5012_Farbteil_BL",
                      B5010_TB5005 := "B5010_TB5005",
                      B5013_TB5006 := "B5013_TB5006",
                      B5014_TB5006 := "B5014_TB5006",
                      B5015_Teil_in_Pos := "B5015_Teil_in_Pos",
                      B5019_TB5009 := "B5019_TB5009",
                      B5021_TB5010 := "B5021_TB5010",
                      B5020_TB5009 := "B5020_TB5009",
                      B5022_TB5010 := "B5022_TB5010",
                      B5016_Teil_vorhanden := "B5016_Teil_vorhanden",
                      xAnlageEin := "100_DB_Kommissionierung".xAnlageEin,
                      xNotAus := "100_DB_Kommissionierung".xNotAusOK,
                      xHauptschalter := "S0_HS",
                      STOP5001 => "STOP5001",
                      STOP5002 => "STOP5002",
                      TB5008 => "TB5008",
                      TB5001 => "TB5001",
                      Emitter_1 => "Emitter_1",
                      TB5002 => "TB5002",
                      TB5003 => "TB5003",
                      TB5004 => "TB5004",
                      TB5005 => "TB5005",
                      STOP5005 => "STOP5005",
                      RS5001_V => "RS5001_V",
                      TB5006 => "TB5006",
                      STOP5003 => "STOP5003",
                      STOP5004 => "STOP5004",
                      TB5007 => "TB5007",
                      RS5001_links => "RS5001_links",
                      TB5009 => "TB5009",
                      TB5010 => "TB5010");
END_REGION

REGION Network 17: Greifarm 4
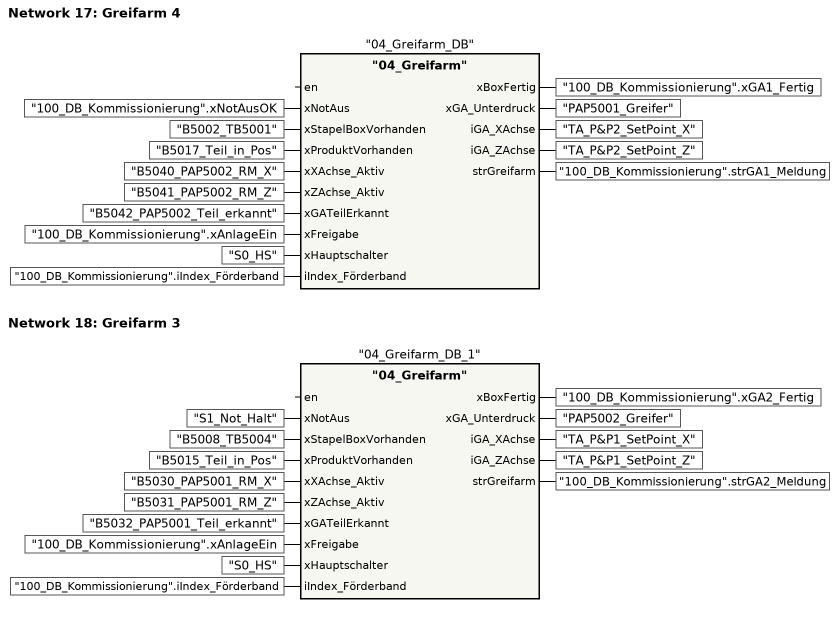
   "04_Greifarm_DB"(xNotAus := "100_DB_Kommissionierung".xNotAusOK,   // "04_Greifarm"
                    xStapelBoxVorhanden := "B5002_TB5001",
                    xProduktVorhanden := "B5017_Teil_in_Pos",
                    xXAchse_Aktiv := "B5040_PAP5002_RM_X",
                    xZAchse_Aktiv := "B5041_PAP5002_RM_Z",
                    xGATeilErkannt := "B5042_PAP5002_Teil_erkannt",
                    xFreigabe := "100_DB_Kommissionierung".xAnlageEin,
                    xHauptschalter := "S0_HS",
                    iIndex_Förderband := "100_DB_Kommissionierung".iIndex_Förderband,
                    xBoxFertig => "100_DB_Kommissionierung".xGA1_Fertig,
                    xGA_Unterdruck => "PAP5001_Greifer",
                    iGA_XAchse => "TA_P&P2_SetPoint_X",
                    iGA_ZAchse => "TA_P&P2_SetPoint_Z",
                    strGreifarm => "100_DB_Kommissionierung".strGA1_Meldung);
END_REGION

REGION Network 18: Greifarm 3
   "04_Greifarm_DB_1"(xNotAus := "S1_Not_Halt",   // "04_Greifarm"
                      xStapelBoxVorhanden := "B5008_TB5004",
                      xProduktVorhanden := "B5015_Teil_in_Pos",
                      xXAchse_Aktiv := "B5030_PAP5001_RM_X",
                      xZAchse_Aktiv := "B5031_PAP5001_RM_Z",
                      xGATeilErkannt := "B5032_PAP5001_Teil_erkannt",
                      xFreigabe := "100_DB_Kommissionierung".xAnlageEin,
                      xHauptschalter := "S0_HS",
                      iIndex_Förderband := "100_DB_Kommissionierung".iIndex_Förderband,
                      xBoxFertig => "100_DB_Kommissionierung".xGA2_Fertig,
                      xGA_Unterdruck => "PAP5002_Greifer",
                      iGA_XAchse => "TA_P&P1_SetPoint_X",
                      iGA_ZAchse => "TA_P&P1_SetPoint_Z",
                      strGreifarm => "100_DB_Kommissionierung".strGA2_Meldung);
END_REGION
END_ORGANIZATION_BLOCK

// folder: Kommissionierung

FUNCTION_BLOCK "03_Förderband"   // FB2, SCL
{ S7_Optimized_Access := 'FALSE' }
VERSION : 0.1
   VAR_INPUT
      B5018_Teil_vorhanden : Bool;
      B5017_Teil_in_Pos : Bool;
      B5002_TB5001 : Bool;
      B5001_TB5001 : Bool;
      xGA1_Fertig : Bool;
      xGA2_Fertig : Bool;
      B5003_TB5002 : Bool;
      B5005_TB5003 : Bool;
      B5004_TB5002 : Bool;
      B5007_TB5004 : Bool;
      B5006_TB5003 : Bool;
      B5009_TB5005 : Bool;
      B5008_TB5004 : Bool;
      B5011_Farbteil_GN : Bool;
      B5012_Farbteil_BL : Bool;
      B5010_TB5005 : Bool;
      B5013_TB5006 : Bool;
      B5014_TB5006 : Bool;
      B5015_Teil_in_Pos : Bool;
      B5019_TB5009 : Bool;
      B5021_TB5010 : Bool;
      B5020_TB5009 : Bool;
      B5022_TB5010 : Bool;
      B5016_Teil_vorhanden : Bool;
      xAnlageEin : Bool;
      xNotAus : Bool;
      xHauptschalter : Bool;
   END_VAR
   VAR_OUTPUT
      STOP5001 : Bool;
      STOP5002 : Bool;
      TB5008 : Bool;
      TB5001 : Bool;
      Emitter_1 : Bool;
      TB5002 : Bool;
      TB5003 : Bool;
      TB5004 : Bool;
      TB5005 : Bool;
      STOP5005 : Bool;
      RS5001_V : Bool;
      TB5006 : Bool;
      STOP5003 : Bool;
      STOP5004 : Bool;
      TB5007 : Bool;
      RS5001_links : Bool;
      TB5009 : Bool;
      TB5010 : Bool;
   END_VAR
   VAR
      stat_iIndex : Int;
      IEC_Timer_0_blau : TON;
      stat_strFörderband : String[15];
      stat_Ntrig1 : Bool;
      stat_Ntig1M : Bool;
      stat_Ntrig2 : Bool;
      stat_Ntig2M : Bool;
      IEC_Timer_1_grün : TON;
   END_VAR
BEGIN
   // ==============================Förderband=======================================
   // Es können zwei verschiedene Produkte über diese Anlage verteilt werden.
   // Blaue oder grüne Produkte.
   // Es darf sich immer nur ein Produkt in der Anlage befinden.

   // Abfrage Hauptschalter
   REGION Abfrage Hauptschalter
       IF NOT #xHauptschalter THEN
           #STOP5001 := 0;
           #STOP5002 := 0;
           #STOP5003 := 0;
           #STOP5004 := 0;
           #STOP5005 := 0;
           #TB5001 := 0;
           #TB5002 := 0;
           #TB5003 := 0;
           #TB5004 := 0;
           #TB5005 := 0;
           #TB5006 := 0;
           #TB5007 := 0;
           #TB5008 := 0;
           #TB5009 := 0;
           #TB5010 := 0;
           #Emitter_1 := 0;
           #RS5001_V := 0;
           #RS5001_links := 0;
           #stat_iIndex := 0;
           #stat_strFörderband := 'HS aus';
           RETURN;
       END_IF;
   END_REGION

   // Abfrage NotAus
   REGION Abfrage NOTAUS
       IF NOT #xNotAus OR "100_DB_Kommissionierung".xAnlageAusgeschaltet THEN
           #STOP5001 := 0;
           #STOP5002 := 0;
           #STOP5003 := 0;
           #STOP5004 := 0;
           #STOP5005 := 0;
           #TB5001 := 0;
           #TB5002 := 0;
           #TB5003 := 0;
           #TB5004 := 0;
           #TB5005 := 0;
           #TB5006 := 0;
           #TB5007 := 0;
           #TB5008 := 0;
           #TB5009 := 0;
           #TB5010 := 0;
           #Emitter_1 := 0;
           #RS5001_V := 0;
           #RS5001_links := 0;
           #stat_iIndex := 0;
           RETURN;
       END_IF;
   END_REGION

   // Entscheidung welches Produkt am Eingang liegt 
   REGION Entscheidung welche Produkt am Eingang liegt
       IF #stat_iIndex = 0 THEN
           #stat_strFörderband := 'Betriebsbereit';
       END_IF;



       IF NOT #B5018_Teil_vorhanden AND #stat_iIndex = 0 AND #xAnlageEin THEN
           #Emitter_1 := 1;
           #STOP5001 := 1;
           #STOP5003 := 1;
           #stat_iIndex := 100;

       END_IF;

       IF NOT #B5016_Teil_vorhanden AND #stat_iIndex = 0 AND #xAnlageEin THEN
           #Emitter_1 := 1;
           #STOP5001 := 1;
           #STOP5003 := 1;
           #stat_iIndex := 200;

       END_IF;
   END_REGION

   // Förderband
   CASE #stat_iIndex OF
       100:    // Stopper ausfahren und Stapelkiste erzeugen
           REGION Stopper ausfahren und Stapelkiste erzeugen

               #STOP5002 := 1;
               #stat_strFörderband := 'In Betrieb';

               // Schritt erhöhen
               IF #B5001_TB5001 THEN
                   #stat_iIndex := #stat_iIndex + 1;
               END_IF;

           END_REGION

       101:    //Förderbänder starten
           REGION Förderbänder starten
               #TB5008 := 1;
               #TB5001 := 1;
               #Emitter_1 := 0;

               IF NOT #B5017_Teil_in_Pos THEN
                   #TB5008 := 0;
               END_IF;


               IF #B5002_TB5001 THEN
                   #TB5001 := 0;
               END_IF; 

               // Zurücksetzen aus vorherigen Schritten
               #Emitter_1 := 0;

               // Schritt erhöhen
               IF NOT #B5017_Teil_in_Pos AND #B5002_TB5001 THEN
                   #stat_iIndex := #stat_iIndex + 1;
               END_IF;
           END_REGION

       102:    // Greifarm abwarten und abtransport über das nächse Förderband
           REGION Greifarm abwarten und abtransport über das nächse Förderband
               IF #xGA1_Fertig THEN
                   (* #STOP5001 := 0; *) // Kann oben bleiben
                   #STOP5002 := 0;
               END_IF;

               IF (* #STOP5001 = 0 AND *) #STOP5002 = 0 THEN
                   #TB5001 := 1;
                   #TB5002 := 1;
               END_IF;

               IF #B5003_TB5002 AND NOT #B5002_TB5001 THEN
                   #TB5001 := 0;
                   #TB5003 := 1;
               END_IF;

               // Schritt erhöhung
               IF NOT #TB5001 AND #TB5002 THEN
                   #stat_iIndex := #stat_iIndex + 1;
               END_IF;
           END_REGION

       103:    // Förderbänder bis zur Farberkennung
           REGION Förderbänder bis zur Farberkennung
               // TB 5002 aus und TB 5003 ein

               IF #B5005_TB5003 AND NOT #B5004_TB5002 THEN
                   #TB5002 := 0;
               END_IF;

               // TB 5003 aus und TB5004 ein
               IF #B5007_TB5004 AND NOT #B5006_TB5003 THEN
                   #TB5003 := 0;
               END_IF;

               IF #B5006_TB5003 THEN
                   #TB5004 := 1;
               END_IF;

               // TB 5004 aus und TB 5005 ein
               IF #B5009_TB5005 AND NOT #B5008_TB5004 THEN
                   #TB5004 := 0;
               END_IF;

               IF #B5008_TB5004 THEN
                   #TB5005 := 1;
               END_IF;

               // Schitt erhöhung
               IF #B5009_TB5005 AND NOT #B5008_TB5004 THEN
                   #stat_iIndex := #stat_iIndex + 1;
               END_IF;

           END_REGION

       104:    // Farberkennung 
           REGION Farberkennung
               // Für blaue Produkte springen wir in 110 
               // Für grüne Produkte springen wir in 210
               IF #B5012_Farbteil_BL THEN
                   #stat_iIndex := 110;
               END_IF;

               IF #B5011_Farbteil_GN THEN
                   #stat_iIndex := 210;
               END_IF;
           END_REGION

       110:    // Rollenförderband blau
           REGION Rollenförderband blau
               #STOP5005 := 1;
               #RS5001_links := 0;
               #RS5001_V := 1;
               #TB5006 := 1;

               IF #B5013_TB5006 AND NOT #B5010_TB5005 THEN
                   #TB5005 := 0;
               END_IF;

               // Flankenauswertung Sensor B5013_TB5006
               // NTrig
               #stat_Ntrig1 := NOT #B5013_TB5006 AND #stat_Ntig1M;
               #stat_Ntig1M := #B5013_TB5006;

               IF #TB5006 = 1 AND #stat_Ntrig1 THEN
                   #STOP5005 := 0;
                   #RS5001_V := 0;
                   #stat_iIndex := #stat_iIndex + 1;
               END_IF;


           END_REGION

       111:    // Remove blaues Produkt 
           REGION Remove blaues Produkt
               #IEC_Timer_0_blau(IN := #B5014_TB5006,
                                     PT := t#0.5s);
                   IF #B5014_TB5006 (* AND #IEC_Timer_0_blau.Q *) THEN
                   #TB5006 := 0;
                   IF NOT #B5015_Teil_in_Pos AND #xAnlageEin THEN
                       #stat_iIndex := 200;
                       #Emitter_1 := 1;
                   ELSE
                       #stat_iIndex := 0;
                   END_IF;
               END_IF;

           END_REGION

       200:    // Stopper ausfahren und Stapelkiste erzeugen
           REGION Stopper ausfahren und Stapelkiste erzeugen

               #STOP5004 := 1;
               #stat_strFörderband := 'In Betrieb';

               // Schritt erhöhen
               IF #B5001_TB5001 THEN
                   #stat_iIndex := #stat_iIndex + 1;
               END_IF;
           END_REGION

       201:    // Förderbänder starten
           REGION Förderbänder starten
               #TB5007 := 1;
               #Emitter_1 := 0;

               IF NOT #B5015_Teil_in_Pos THEN
                   #TB5007 := 0;
               END_IF;

               // TB5001
               IF #B5001_TB5001 THEN
                   #TB5001 := 1;
               END_IF;

               IF #B5003_TB5002 AND NOT #B5002_TB5001 THEN
                   #TB5001 := 0;
               END_IF;

               // TB 5002
               IF #B5002_TB5001 THEN
                   #TB5002 := 1;
               END_IF;

               IF #B5005_TB5003 AND NOT #B5004_TB5002 THEN
                   #TB5002 := 0;
               END_IF;

               // TB 5003
               IF #B5004_TB5002 THEN
                   #TB5003 := 1;
               END_IF;

               IF #B5007_TB5004 AND NOT #B5006_TB5003 THEN
                   #TB5003 := 0;
               END_IF;

               // TB 5004
               IF #B5006_TB5003 THEN
                   #TB5004 := 1;
               END_IF;

               IF #B5008_TB5004 THEN
                   #TB5004 := 0;
               END_IF;

               // Schitt erhöhung
               IF #B5008_TB5004 THEN
                   #stat_iIndex := #stat_iIndex + 1;
               END_IF;

           END_REGION

       202:    // Greifarm abwarten und abtransport über das nächse Förderband
           REGION Greifarm abwarten und abtransport über das nächse Förderband
               IF #xGA2_Fertig THEN
                   (* #STOP5003 := 0; *) // Kann oben bleiben
                   #STOP5004 := 0;
               END_IF;

               IF (* #STOP5003 = 0 AND *) #STOP5004 = 0 THEN
                   #TB5004 := 1;
                   #TB5005 := 1;
               END_IF;

               IF #B5009_TB5005 AND NOT #B5008_TB5004 THEN
                   #TB5004 := 0;
               END_IF;

               // Schritt erhöhung
               IF #B5009_TB5005 AND NOT #B5008_TB5004 THEN
                   #stat_iIndex := #stat_iIndex + 1;
               END_IF;
           END_REGION

       203:    // Farberkennung
           REGION Farberkennung
               // Für blaue Produkte springen wir in 110 
               // Für grüne Produkte springen wir in 210
               IF #B5012_Farbteil_BL THEN
                   #stat_iIndex := 110;
               END_IF;

               IF #B5011_Farbteil_GN THEN
                   #stat_iIndex := 210;
               END_IF;
           END_REGION

       210:    //Rollenförderband grün
           REGION Rollenförderband grün
               #STOP5005 := 1;
               #RS5001_V := 1;
               #RS5001_links := 1;
               #TB5009 := 1;

               IF #B5019_TB5009 AND NOT #B5010_TB5005 THEN
                   #TB5005 := 0;
               END_IF;

               // Flankenauswertung Sensor B5013_TB5006
               // NTrig
               #stat_Ntrig2 := NOT #B5019_TB5009 AND #stat_Ntig2M;
               #stat_Ntig2M := #B5019_TB5009;

               IF #TB5009 = 1 AND #stat_Ntrig2 THEN
                   #STOP5005 := 0;
                   #RS5001_V := 0;
                   #stat_iIndex := #stat_iIndex + 1;
               END_IF;


           END_REGION

       211:    // Remove grünes Produkt
           REGION Remove grünes Produkt

               // TB 5009
               IF #B5021_TB5010 AND NOT #B5020_TB5009 THEN
                   #TB5009 := 0;
               END_IF;

               // TB 5010   
               IF #B5020_TB5009 THEN
                   #TB5010 := 1;
               END_IF;

               #IEC_Timer_1_grün(IN := #B5022_TB5010,
                                 PT := t#0.5s);


               IF #B5022_TB5010 (* AND NOT #IEC_Timer_1_grün.Q *) THEN
                   #TB5010 := 0;
                   IF NOT #B5017_Teil_in_Pos AND #xAnlageEin THEN
                       #stat_iIndex := 100;
                       #Emitter_1 := 1;
                   ELSE
                       #stat_iIndex := 0;
                   END_IF;
               END_IF;

               END_REGION


       ELSE  // Error
           #stat_strFörderband := 'Error';
           ;
   END_CASE;

   // Schrittangabe
   "100_DB_Kommissionierung".iIndex_Förderband := #stat_iIndex;
END_FUNCTION_BLOCK

FUNCTION_BLOCK "04_Greifarm"   // FB3, SCL
{ S7_Optimized_Access := 'FALSE' }
VERSION : 0.1
   VAR_INPUT
      xNotAus : Bool;
      xStapelBoxVorhanden : Bool;
      xProduktVorhanden : Bool;
      xXAchse_Aktiv : Bool;
      xZAchse_Aktiv : Bool;
      xGATeilErkannt : Bool;
      xFreigabe : Bool;
      xHauptschalter : Bool;
      iIndex_Förderband : Int;
   END_VAR
   VAR_OUTPUT
      xBoxFertig : Bool;
      xGA_Unterdruck : Bool;
      iGA_XAchse : Int;
      iGA_ZAchse : Int;
      strGreifarm : String[30];
   END_VAR
   VAR
      stat_iSchritt : Int;
      stat_strGA : String[30];
      xNtrig_XAchse : Bool;
      xNtrig_XAchseM : Bool;
      xNtrig_ZAchse : Bool;
      xNtrig_ZAchseM : Bool;
      stat_rGA_XAchse : Real;
      stat_rGA_ZAchse : Real;
      stat_rPos_Ga_XAchse : Real;
      stat_rPos_GA_ZAchse : Real;
   END_VAR
   VAR_TEMP
      temp_ErrorGA_XAchse : Word;
      temp_ErrorGA_ZAchse : Word;
      temp_Ret_Val_XAchse : Word;
      temp_Ret_Val_ZAchse : Word;
   END_VAR
BEGIN
   // ======================== Greifarm =====================
   // Der Greifarm soll grüne oder blaue Produkte in eine Stapelbox legen

   // Startbedingung
   REGION Startbedingung
       // xProduktVorhanden kommt von der Lichtschranke (0 = Produkt da, 1 = kein Produkt da)
       IF #xStapelBoxVorhanden AND NOT #xProduktVorhanden AND #stat_iSchritt = 0
           AND #xFreigabe AND (#iIndex_Förderband = 102 OR #iIndex_Förderband = 202) (* AND NOT #xXAchse_Pos AND NOT #xZAchse_Pos *)THEN
           #stat_iSchritt := 1;
       END_IF;
   END_REGION

   // Flankenauswertung
   REGION Flankenauswertung
       // Flankenauswertung für X Achse (NTrig)
       #xNtrig_XAchse := NOT #xXAchse_Aktiv AND #xNtrig_XAchseM;
       #xNtrig_XAchseM := #xXAchse_Aktiv;

       // Flankenauswertung für Z Achse (NTrig)
       #xNtrig_ZAchse := NOT #xZAchse_Aktiv AND #xNtrig_ZAchseM;
       #xNtrig_ZAchseM := #xZAchse_Aktiv;
   END_REGION

   // Sacle PosX & PosZ => wird nicht verwendet mangels Analogeingänge
   REGION Sacle PosX & PosZ 
       (* #temp_Ret_Val_XAchse := SCALE(IN := #iXAchse_Pos, HI_LIM := 10.0, LO_LIM := 0.0, BIPOLAR := False, OUT => #stat_rPos_Ga_XAchse);

       #temp_Ret_Val_ZAchse := SCALE(IN := #iZAchse_Pos, HI_LIM := 10.0, LO_LIM := 0.0, BIPOLAR := False, OUT => #stat_rPos_GA_ZAchse); *)
   END_REGION

   // Unscale für X & Z Achse
   REGION Unscale und Convert für X & Z Achse
       // X-Achse
       // Unscale r=>i und dann Convert i=>w
       #temp_ErrorGA_XAchse := UNSCALE(IN := #stat_rGA_XAchse, HI_LIM := 10.0, LO_LIM := 0.0, BIPOLAR := false, OUT => #iGA_XAchse);


       // Y-Achse
       // Unscale r=>i und dann Convert i=>w
       #temp_ErrorGA_ZAchse := UNSCALE(IN := #stat_rGA_ZAchse, HI_LIM := 10.0, LO_LIM := 0.0, BIPOLAR := false, OUT => #iGA_ZAchse);

   END_REGION

   // Schrittkette Greifarm
   REGION Schrittkette
       CASE #stat_iSchritt OF

           0:  // Ruhezustand
               REGION Schritt 0 Ruhezustand
                   #stat_strGA := 'Betriebsbereit';
                   #stat_rGA_XAchse := 0.0;
                   #stat_rGA_ZAchse := 0.0;
               END_REGION

           1:  // Schritt 1: X Achse ausfahren auf 6.7
               REGION Schritt 1 X Achse ausfahren
                   #stat_rGA_XAchse := 6.7;
                   #stat_strGA := 'X Achse ausfahren';

                   // Schritt erhöhen
                   IF #xNtrig_XAchse = 1 THEN
                       #stat_iSchritt := 2;
                   END_IF;
               END_REGION

           2:  // Schritt 2: Z Achse ausfahren
               REGION Schritt 2 Z Achse ausfahren
                   #stat_rGA_ZAchse := 10.0;
                   #stat_strGA := 'Z Achse ausfahren';

                   // Schritt erhöhen
                   IF #xNtrig_ZAchse = 1 THEN
                       #stat_iSchritt := 3;
                   END_IF;
               END_REGION

           3:  // Schritt 3: Teil Erkennung und Unterdruck Erzeugung
               REGION Schritt 3 Unterdruck erzeugen
                   #xGA_Unterdruck := 1;
                   #stat_strGA := 'Unterdruck an, Teil erkennen';

                   // Schritt erhöhen
                   IF #xGATeilErkannt THEN
                       #stat_iSchritt := 4;
                   END_IF;
               END_REGION

           4:  // Schritt 4: Z Achse einfahren
               REGION Schritt 4 Z Achse einfahren
                   #stat_rGA_ZAchse := 0.0;
                   #stat_strGA := 'Z Achse einfahren';

                   // Schritt erhöhen
                   IF #xNtrig_ZAchse = 1 THEN
                       #stat_iSchritt := 5;
                   END_IF;
               END_REGION

           5:  // Schritt 5: X Achse einfahren
               REGION Schritt 5 X Achse einfahren
                   #stat_rGA_XAchse := 0.0;
                   #stat_strGA := 'X Achse einfahren';

                   // Schritt erhöhen
                   IF #xNtrig_XAchse = 1 THEN
                       #stat_iSchritt := 6;
                   END_IF;
               END_REGION

           6:  // Schritt 6: Z Achse ausfahren
               REGION Schritt 6 Z Achse ausfahren
                   #stat_rGA_ZAchse := 10.0;
                   #stat_strGA := 'Z Achse Ausfahren';

                   // Schritt erhöhen
                   IF #xNtrig_ZAchse = 1 THEN
                       #stat_iSchritt := 7;
                   END_IF;
               END_REGION

           7:  // Schritt 7: Unterdruck beenden
               REGION Schritt 7 Unterdruck beenden
                   #xGA_Unterdruck := 0;

                   // Schritt erhöhen
                   #stat_iSchritt := 8;
               END_REGION

           8:  // Schritt 8: Z Achse einfahren
               REGION Schritt 8 Z Achse einfahren
                   #stat_rGA_ZAchse := 0.0;
                   #stat_strGA := 'Z Achse Einfahren';

                   // Schritt erhöhen
                   IF #xNtrig_ZAchse = 1 THEN
                       #stat_iSchritt := 9;
                   END_IF;
               END_REGION

           9:  // Schritt 9: Box fertig, warten bis die Box weg ist
               REGION Schritt 9 Box fertig
                   #stat_strGA := 'Box fertig';

                   IF NOT #xStapelBoxVorhanden THEN
                       #stat_iSchritt := 0;
                   END_IF;
               END_REGION

           ELSE  // Error
               #stat_strGA := 'ERROR';
               #stat_iSchritt := 0;

       END_CASE;
   END_REGION

   // Meldung für die Bandsteuerung
   REGION Meldung Box fertig
       #xBoxFertig := #stat_iSchritt = 9;
       #strGreifarm BLKMOV #stat_strGA;
   END_REGION

   // Abfrage Hauptschalter
   REGION Abfrage Hauptschalter
       IF NOT #xHauptschalter THEN
           #stat_iSchritt := 0;
           #iGA_XAchse := 0;
           #iGA_ZAchse := 0;
           #xGA_Unterdruck := 0;
           #xBoxFertig := 0;
           #stat_strGA := 'Hauptschalter aus';
       END_IF;
   END_REGION

   // Abfrage NotAus
   REGION Abfrage NOTAUS
       IF NOT #xNotAus THEN
           #stat_iSchritt := 0;
           #iGA_XAchse := 0;
           #iGA_ZAchse := 0;
           #xGA_Unterdruck := 0;
           #xBoxFertig := 0;
           #stat_strGA := 'NOT-AUS';
       END_IF;
   END_REGION
END_FUNCTION_BLOCK

FUNCTION_BLOCK "02_AnlageEinAus"   // FB9, SCL
{ S7_Optimized_Access := 'FALSE' }
VERSION : 0.1
   VAR_INPUT
      xHauptschalter : Bool;
      xEinTaster : Bool;
      xNotAusDB : Bool;
      xAusTaster : Bool;
      xBlinklichttakt : Bool;
   END_VAR
   VAR_OUTPUT
      xSirene : Bool;
      xRundumleuchte : Bool;
      xMS_Grün : Bool;
      xMS_Gelb : Bool;
      xMS_Rot : Bool;
      xMT_Grün : Bool;
      xMT_Rot : Bool;
      xAnlageStartet : Bool;
      xAnlageEin : Bool;
      xAnlageAusgeschaltet : Bool;
   END_VAR
   VAR
      IEC_Timer_0_AnlageEinAus : TON;
      stat_xAnlageAusgeschaltet : Bool;
      stat_xAnlageStartet : Bool;
      stat_xAnlageEin : Bool;
   END_VAR
BEGIN
   //==============================Beschreibung======================================
   // -Damit die Anlage starten kann muss der Hauptschalter eingeschalten und der Starttaster betätigt werden
   // -Zusätzlich muss die NotAus Bedingung ein Highsignal führen
   // -Wird der Stopptaster betätigt, wird der aktuelle Vorgang abgeschlossen und nicht erneut gestartet
   // -Der Anlagenstart wird über die Sirene und Rundumleuchte für 10s nach betätigen des Starttasters gemeldet
   //  erst nach ablauf der 10s fährt die Anlage an
   // -Die Meldeleuchten geben die aktuelle Betriebsart an

   // Abfrage Hauptschalter
    REGION Abfrage Hauptschalter
        IF NOT #xHauptschalter THEN
            #stat_xAnlageStartet := 0;
            #stat_xAnlageEin := 0;
            #xSirene := 0;
            #xRundumleuchte := 0;
            #xMS_Grün := 0;
            #xMS_Gelb := 0;
            #xMS_Rot := 0;
            #xMT_Grün := 0;
            #xMT_Rot := 0;
            #stat_xAnlageAusgeschaltet := 0;
            RETURN;
        END_IF;
    END_REGION

   // ============Abfrage NotAus=======
    REGION Abfrage NotAus
        IF NOT #xNotAusDB THEN
            #stat_xAnlageStartet := 0;
            #stat_xAnlageEin := 0;
            #xSirene := 0;
            #xRundumleuchte := 0;
            #xMS_Grün := 0;
            #xMS_Gelb := 0;
            #xMS_Rot := 1 AND "Takt_1HZ";
            #xMT_Grün := 0;
            #xMT_Rot := 0;
            #stat_xAnlageAusgeschaltet := 0;
            RETURN;
        END_IF;
    END_REGION


   // ============Anlage Ein===========
   REGION Anlage Ein
       IF  #xEinTaster AND NOT #stat_xAnlageStartet AND NOT #stat_xAnlageEin THEN
           #stat_xAnlageStartet := 1;
           ;
       END_IF;


       IF #IEC_Timer_0_AnlageEinAus.Q THEN
           #stat_xAnlageStartet := 0;
           #stat_xAnlageEin := 1;
       END_IF;
   END_REGION

   // ============Anlage Aus===========
   REGION Anlage Aus    
       IF NOT #xAusTaster THEN
           #stat_xAnlageStartet := 0;
           #stat_xAnlageEin := 0;
       END_IF;

   END_REGION

   // ============Signale==============
   REGION Signale
       // Sirene und Rundumleuchte
       REGION SireneRundumleuchte
           IF NOT #IEC_Timer_0_AnlageEinAus.Q AND #stat_xAnlageStartet THEN
               #xSirene := 1;
               #xRundumleuchte := 1;
           ELSE
               #xSirene := 0;
               #xRundumleuchte := 0;
           END_IF;
       END_REGION

       // Anlage Inbetrieb
       REGION AnlageInbetrieb
           IF #stat_xAnlageStartet OR #stat_xAnlageEin THEN
               #xMS_Grün := 1;
               #xMT_Grün := 1;
           ELSE
               #xMS_Grün := 0;
               #xMT_Grün := 0;
           END_IF;
       END_REGION

       // Anlage Betriebsbereit
       REGION AnlageInbetrieb
           IF #xHauptschalter AND #xBlinklichttakt AND NOT #stat_xAnlageStartet AND NOT #stat_xAnlageEin AND NOT #stat_xAnlageAusgeschaltet THEN
               #xMS_Gelb := 1;
           ELSE
               #xMS_Gelb := 0;
           END_IF;
       END_REGION

           // Anlage Aus
       REGION AnlageAus

           IF NOT #xAusTaster AND (#xHauptschalter OR #xNotAusDB) THEN
               #stat_xAnlageAusgeschaltet := 1;
               #xMT_Rot := 1;
           END_IF;

           IF #xEinTaster THEN
               #stat_xAnlageAusgeschaltet := 0;
               #xMT_Rot := 0;
           END_IF;

           #xMS_Rot := #stat_xAnlageAusgeschaltet AND #xBlinklichttakt;

       END_REGION

   END_REGION

   // ============Zeitfunktionen=======
   #IEC_Timer_0_AnlageEinAus(IN:=#stat_xAnlageStartet,
                             PT:=t#10s);

   // ============Static zu Output=====
   #xAnlageStartet := #stat_xAnlageStartet;
   #xAnlageEin := #stat_xAnlageEin;
   #xAnlageAusgeschaltet := #stat_xAnlageAusgeschaltet;
END_FUNCTION_BLOCK

FUNCTION "01_NotAus_STO" : Void   // FC1, SCL
{ S7_Optimized_Access := 'FALSE' }
VERSION : 0.1
   VAR_INPUT
      xNotAus : Bool;
   END_VAR
   VAR_OUTPUT
      xNotAusOK : Bool;
   END_VAR
BEGIN
   //==============================NotAus======================================
   //STO Energiezufuhr wird sofort abgeschaltet wenn der NotAus betätigt wird
   //Der NotAus ist als Öffner-Kontakt ausgeführt => Drahtbruchsicher


   IF #xNotAus THEN
       #xNotAusOK:= 1
       ;
   END_IF;
END_FUNCTION

// folder: Montage/Bearbeitung Blau

FUNCTION_BLOCK "01Transportband vor Bearbeitung"   // FB1, FBD
{ S7_Optimized_Access := 'FALSE' }
VERSION : 0.1
   VAR_TEMP   // added for the SCL form of the ladder/FBD networks
      _w1 : Bool;
   END_VAR
BEGIN

REGION Network 1: "TB3008"
   // Prüft Start/Stop bedingungen 
   // Band 3008 Start nachdem Sensor "B3013_TB3008" unterbrochen wird.
   // Stoppt wenn Sensor "B3011_TB3007" unterbrochen wird.
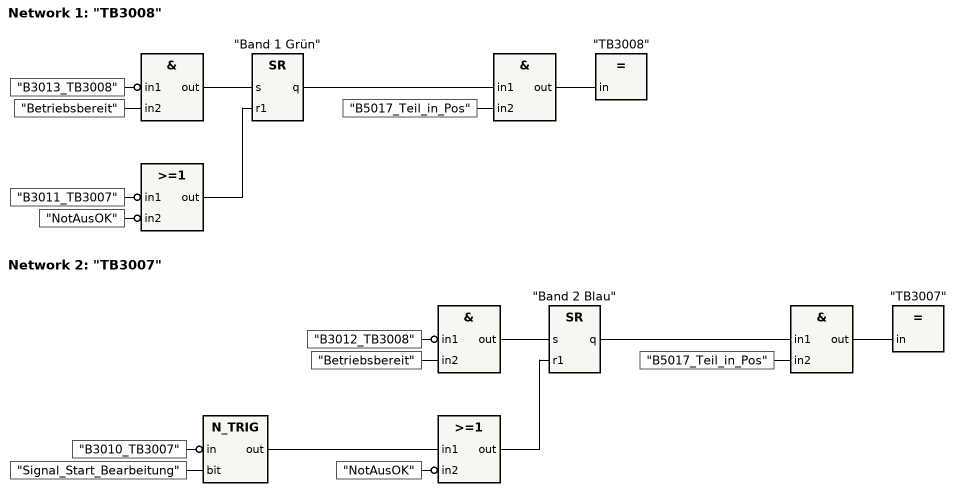
   IF NOT "B3013_TB3008" AND "Betriebsbereit" THEN
       "Band 1 Grün" := TRUE;   // SR flip-flop
   END_IF;
   IF NOT "B3011_TB3007" OR NOT "NotAusOK" THEN "Band 1 Grün" := FALSE; END_IF;
   "TB3008" := "Band 1 Grün" AND "B5017_Teil_in_Pos";
END_REGION

REGION Network 2: "TB3007"
   // Band 3007 Start nachem Sensor "B3012_TB3008" unterbrochen wird.
   // Fällt ab wenn Sensor "B3010_TB3007" unterbrochen wird.
   // Sensor "B3010_TB3007" erzeugt ein Signal für die Weiterverarbeitung:"Signal_Start_Bearbeitung"
   // Prüft Start/Stop bedingungen
   #_w1 := NOT (NOT "B3010_TB3007") AND "Signal_Start_Bearbeitung";   // falling edge
   "Signal_Start_Bearbeitung" := NOT "B3010_TB3007";
   IF NOT "B3012_TB3008" AND "Betriebsbereit" THEN
       "Band 2 Blau" := TRUE;   // SR flip-flop
   END_IF;
   IF #_w1 OR NOT "NotAusOK" THEN "Band 2 Blau" := FALSE; END_IF;
   "TB3007" := "Band 2 Blau" AND "B5017_Teil_in_Pos";
END_REGION
END_FUNCTION_BLOCK

FUNCTION_BLOCK "03_Weiterverarbeitung"   // FB4, FBD
{ S7_Optimized_Access := 'FALSE' }
VERSION : 0.1
   VAR_TEMP   // added for the SCL form of the ladder/FBD networks
      _w1 : Bool;
   END_VAR
BEGIN

REGION Network 1: "TB3006"
   // Band 3006 Start wenn Sensor "B3009_TB3006" unterbrochen wird.
   // Stoppt wenn Sensor "B3004_TB3001" oder "B3014_TB3005" unterbrochen wird.
   // Prüft Start/Stop bedingungen.
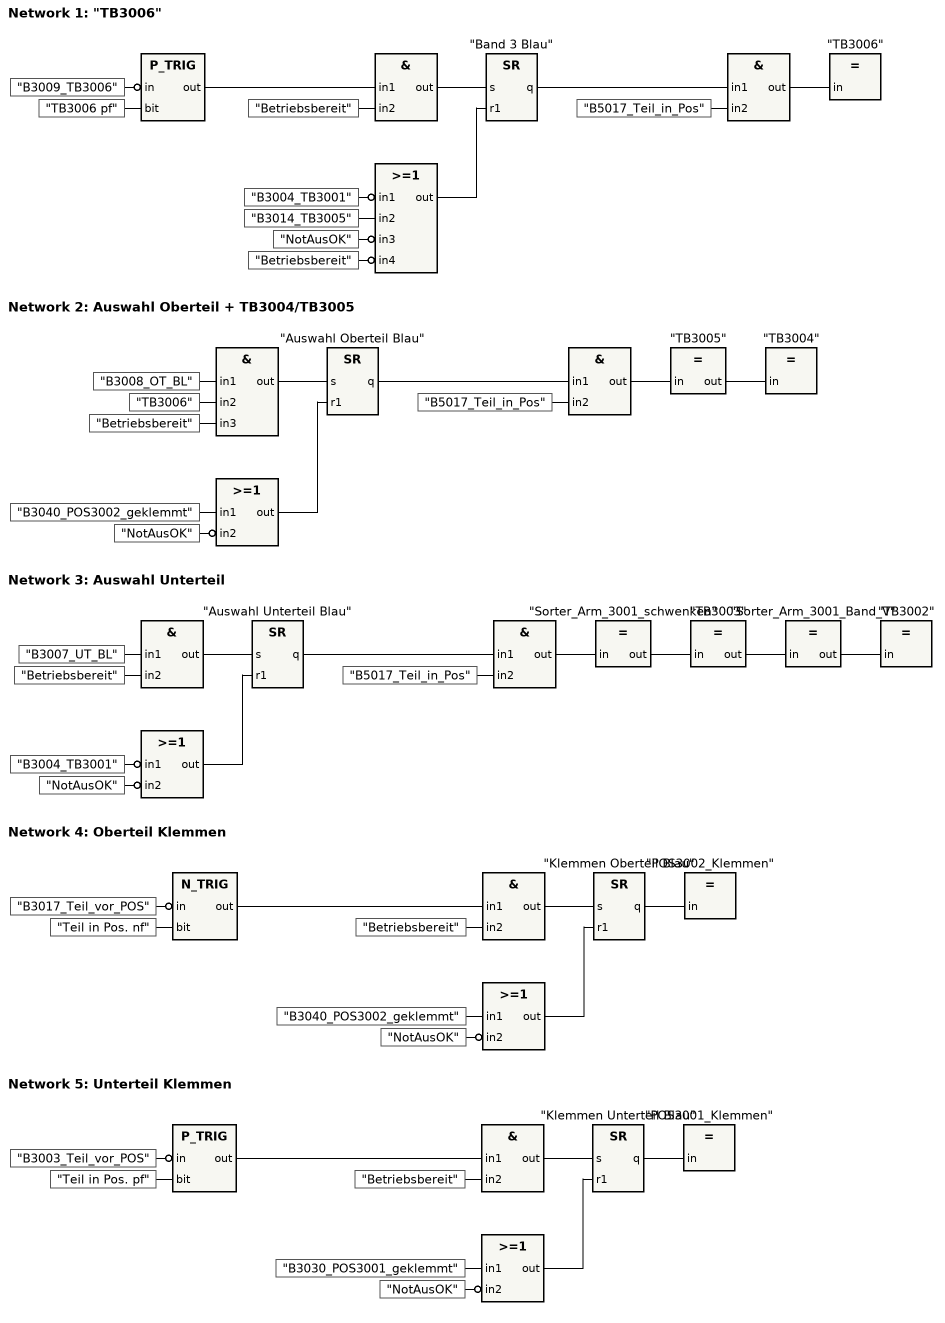
   #_w1 := NOT "B3009_TB3006" AND NOT "TB3006 pf";   // rising edge
   "TB3006 pf" := NOT "B3009_TB3006";
   IF #_w1 AND "Betriebsbereit" THEN
       "Band 3 Blau" := TRUE;   // SR flip-flop
   END_IF;
   IF NOT "B3004_TB3001" OR "B3014_TB3005" OR NOT "NotAusOK" OR NOT "Betriebsbereit" THEN
       "Band 3 Blau" := FALSE;
   END_IF;
   "TB3006" := "Band 3 Blau" AND "B5017_Teil_in_Pos";
END_REGION

REGION Network 2: Auswahl Oberteil + TB3004/TB3005
   // Band "TB3005" und "TB3004" starten wenn der Sensor "B3008_OT_BL" und das Band "TB3006" aktiv ist.
   // Setzt sich zurück sobald Objekt geklemmt wurde mit dem Sensor "B3040_POS3002_geklemmt".
   // Prüft Start/Stop bedingungen.
   IF "B3008_OT_BL" AND "TB3006" AND "Betriebsbereit" THEN
       "Auswahl Oberteil Blau" := TRUE;   // SR flip-flop
   END_IF;
   IF "B3040_POS3002_geklemmt" OR NOT "NotAusOK" THEN "Auswahl Oberteil Blau" := FALSE; END_IF;
   "TB3005" := "Auswahl Oberteil Blau" AND "B5017_Teil_in_Pos";
   "TB3004" := "TB3005";
END_REGION

REGION Network 3: Auswahl Unterteil
   // "Sorter_Arm_3001_schwenken","TB3003","Sorter_Arm_3001_Band_V","TB3002" werden aktiv sobald 
   // Sensor "B3007_UT_BL" reagiert.
   // Setzt sich zurück sobald das Objekt den Sensor "B3004_TB3001" unterbricht.
   // Prüft Start/Stop bedingungen.
   IF "B3007_UT_BL" AND "Betriebsbereit" THEN
       "Auswahl Unterteil Blau" := TRUE;   // SR flip-flop
   END_IF;
   IF NOT "B3004_TB3001" OR NOT "NotAusOK" THEN "Auswahl Unterteil Blau" := FALSE; END_IF;
   "Sorter_Arm_3001_schwenken" := "Auswahl Unterteil Blau" AND "B5017_Teil_in_Pos";
   "TB3003" := "Sorter_Arm_3001_schwenken";
   "Sorter_Arm_3001_Band_V" := "Sorter_Arm_3001_schwenken";
   "TB3002" := "Sorter_Arm_3001_schwenken";
END_REGION

REGION Network 4: Oberteil Klemmen
   // Objekt wird geklemmt sobald es den Sensor "B3017_Teil_vor_POS" unterbricht.
   // Fällt ab sobald Objekt geklemmt wurde: "B3040_POS3002_geklemmt".
   // Prüft Start/Stop bedingungen.
   #_w1 := NOT (NOT "B3017_Teil_vor_POS") AND "Teil in Pos. nf";   // falling edge
   "Teil in Pos. nf" := NOT "B3017_Teil_vor_POS";
   IF #_w1 AND "Betriebsbereit" THEN
       "Klemmen Oberteil Blau" := TRUE;   // SR flip-flop
   END_IF;
   IF "B3040_POS3002_geklemmt" OR NOT "NotAusOK" THEN "Klemmen Oberteil Blau" := FALSE; END_IF;
   "POS3002_Klemmen" := "Klemmen Oberteil Blau";
END_REGION

REGION Network 5: Unterteil Klemmen
   // Objekt wird geklemmt sobald es den Sensor "B3003_Teil_vor_POS" unterbricht.
   // Fällt ab sobald Objekt geklemmt wurde:"B3030_POS3001_geklemmt".
   // Prüft Start/Stop bedingungen.
   #_w1 := NOT "B3003_Teil_vor_POS" AND NOT "Teil in Pos. pf";   // rising edge
   "Teil in Pos. pf" := NOT "B3003_Teil_vor_POS";
   IF #_w1 AND "Betriebsbereit" THEN
       "Klemmen Unterteil Blau" := TRUE;   // SR flip-flop
   END_IF;
   IF "B3030_POS3001_geklemmt" OR NOT "NotAusOK" THEN "Klemmen Unterteil Blau" := FALSE; END_IF;
   "POS3001_Klemmen" := "Klemmen Unterteil Blau";
END_REGION

REGION Network 6: Unterteil TB3001 bis zur Klemme
   // Wenn Sensor "B3005_TB3002" unterbrochen wird oder das Signal "FreigabeKommissionierung" aktiviert sich "TB3001".
   // Fällt ab wenn das Objekt geklemmt wurde.
   // Prüft Start/Stop bedingungen.
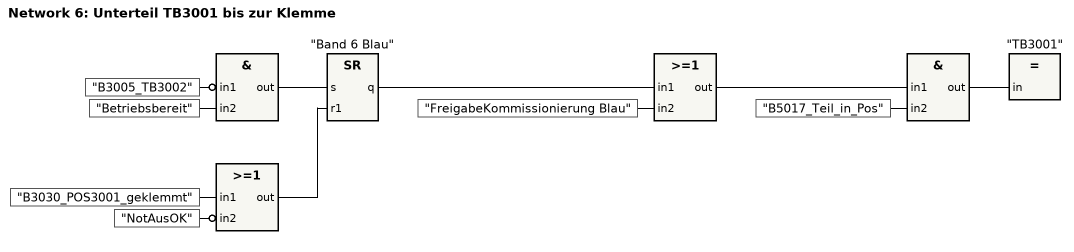
   IF NOT "B3005_TB3002" AND "Betriebsbereit" THEN
       "Band 6 Blau" := TRUE;   // SR flip-flop
   END_IF;
   IF "B3030_POS3001_geklemmt" OR NOT "NotAusOK" THEN "Band 6 Blau" := FALSE; END_IF;
   "TB3001" := ("Band 6 Blau" OR "FreigabeKommissionierung Blau") AND "B5017_Teil_in_Pos";
END_REGION
END_FUNCTION_BLOCK

FUNCTION_BLOCK "04_Zusammenbau"   // FB5, FBD
{ S7_Optimized_Access := 'FALSE' }
VERSION : 0.1
   VAR_TEMP   // added for the SCL form of the ladder/FBD networks
      _w1 : Bool;
      _w2 : Bool;
      _w3 : Bool;
   END_VAR
BEGIN

REGION Network 1: Prüfung Unterteil vorhanden
   // Merker "Freigabe_Zusammenbau UT" wird gesetzt wenn das Objekt geklemmt wurde."POS3001_Klemmen"
   // Fällt ab sobald das fertige Objekt in die Kommissionierung weiter gegeben wurde."B3001_TB3001"
   // Prüft Start/Stop bedingungen.
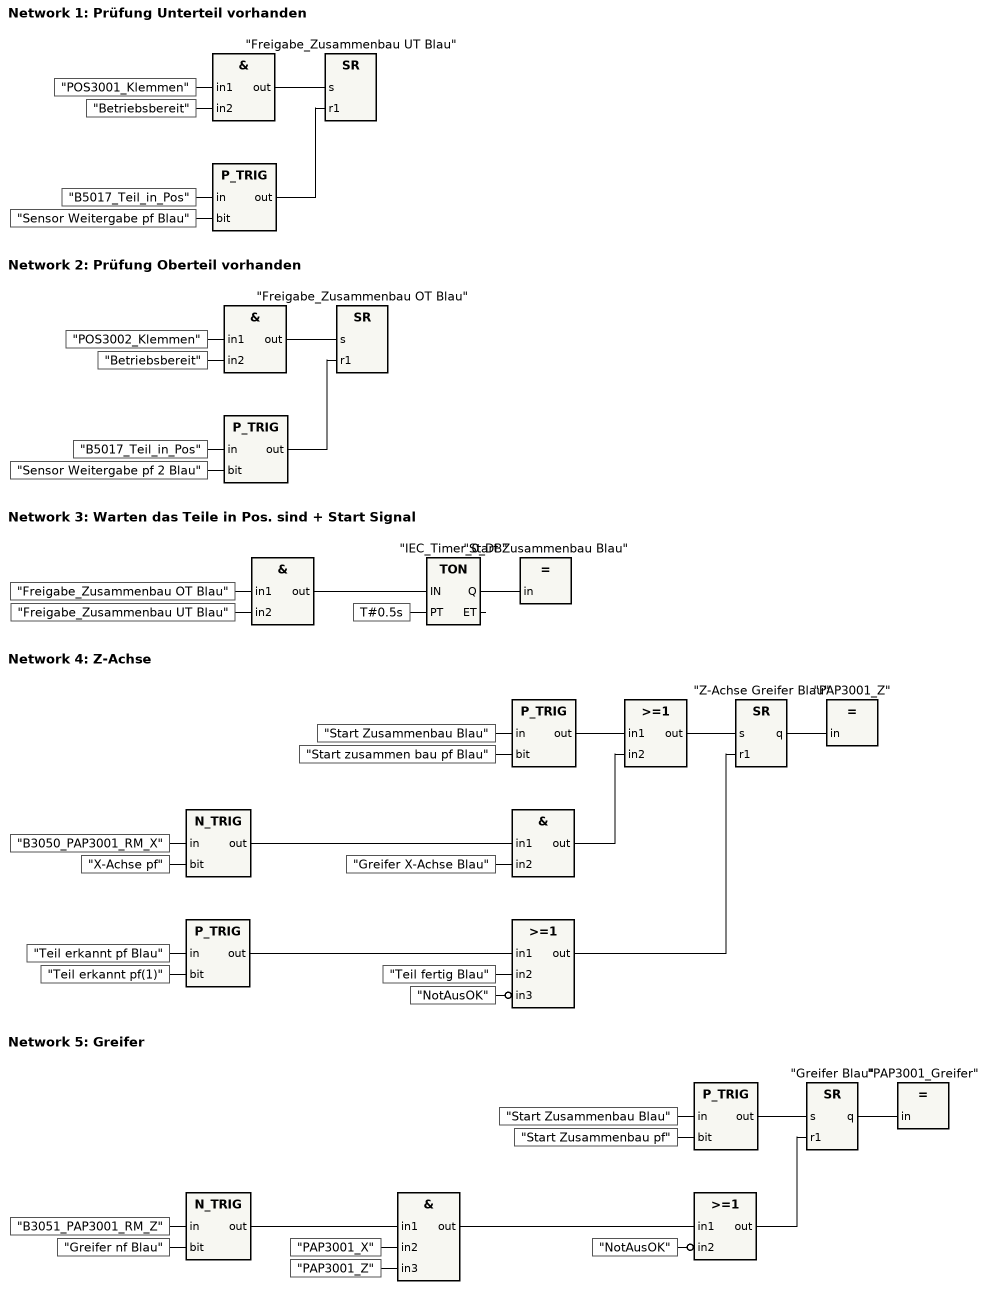
   #_w1 := "B5017_Teil_in_Pos" AND NOT "Sensor Weitergabe pf Blau";   // rising edge
   "Sensor Weitergabe pf Blau" := "B5017_Teil_in_Pos";
   IF "POS3001_Klemmen" AND "Betriebsbereit" THEN
       "Freigabe_Zusammenbau UT Blau" := TRUE;   // SR flip-flop
   END_IF;
   IF #_w1 THEN "Freigabe_Zusammenbau UT Blau" := FALSE; END_IF;
END_REGION

REGION Network 2: Prüfung Oberteil vorhanden
   // Merker"Freigabe_Zusammenbau OT" wird gesetzt wenn das Objekt geklemmt wurde."POS3002_Klemmen"
   // Fällt ab sobald das fertige Objekt in die Kommissionierung weiter gegeben wurde."B3001_TB3001"
   // Prüft Start/Stop bedingungen.
   #_w1 := "B5017_Teil_in_Pos" AND NOT "Sensor Weitergabe pf 2 Blau";   // rising edge
   "Sensor Weitergabe pf 2 Blau" := "B5017_Teil_in_Pos";
   IF "POS3002_Klemmen" AND "Betriebsbereit" THEN
       "Freigabe_Zusammenbau OT Blau" := TRUE;   // SR flip-flop
   END_IF;
   IF #_w1 THEN "Freigabe_Zusammenbau OT Blau" := FALSE; END_IF;
END_REGION

REGION Network 3: Warten das Teile in Pos. sind + Start Signal
   // Sobald beide Freigaben erteilt wurden, wird nach T#0.5s das Signal "Start Zusammenbau" erzeugt.
   "IEC_Timer_0_DB".TON(IN := "Freigabe_Zusammenbau OT Blau" AND "Freigabe_Zusammenbau UT Blau", PT := T#0.5s);
   "Start Zusammenbau Blau" := "IEC_Timer_0_DB".Q;
END_REGION

REGION Network 4: Z-Achse
   // Z-Achse senkt sich sobald das Startsignal "Start Zusammenbau" aktiv ist.
   // Fähr hoch wenn ein Teil erkannt wurde "Teil erkannt pf"oder das das Signal "Teil fertig" kommt.
   // Prüft Start/Stop bedingungen.
   #_w1 := "Start Zusammenbau Blau" AND NOT "Start zusammen bau pf Blau";   // rising edge
   "Start zusammen bau pf Blau" := "Start Zusammenbau Blau";
   #_w2 := NOT "B3050_PAP3001_RM_X" AND "X-Achse pf";   // falling edge
   "X-Achse pf" := "B3050_PAP3001_RM_X";
   #_w3 := "Teil erkannt pf Blau" AND NOT "Teil erkannt pf(1)";   // rising edge
   "Teil erkannt pf(1)" := "Teil erkannt pf Blau";
   IF #_w1 OR (#_w2 AND "Greifer X-Achse Blau") THEN
       "Z-Achse Greifer Blau" := TRUE;   // SR flip-flop
   END_IF;
   IF #_w3 OR "Teil fertig Blau" OR NOT "NotAusOK" THEN "Z-Achse Greifer Blau" := FALSE; END_IF;
   "PAP3001_Z" := "Z-Achse Greifer Blau";
END_REGION

REGION Network 5: Greifer
   // Greifer wird aktiviert sobald das Signal "Start Zusammenbau"kommt.
   // Fällt ab sobald das Objekt fertig zusammen gebaut ist über das Signal "B3051_PAP3001_RM_Z" wenn die jeweiligen X und Z Achsenposition
   // des Roboterarms entsprechend positioniert sind."PAP3001_X","PAP3001_Z".
   // Prüft Stop bedingung.
   #_w1 := "Start Zusammenbau Blau" AND NOT "Start Zusammenbau pf";   // rising edge
   "Start Zusammenbau pf" := "Start Zusammenbau Blau";
   #_w2 := NOT "B3051_PAP3001_RM_Z" AND "Greifer nf Blau";   // falling edge
   "Greifer nf Blau" := "B3051_PAP3001_RM_Z";
   IF #_w1 THEN
       "Greifer Blau" := TRUE;   // SR flip-flop
   END_IF;
   IF (#_w2 AND "PAP3001_X" AND "PAP3001_Z") OR NOT "NotAusOK" THEN "Greifer Blau" := FALSE; END_IF;
   "PAP3001_Greifer" := "Greifer Blau";
END_REGION

REGION Network 6: X-Achse
   // Z-Achse fährt aus sobald ein Teil erkannt wurde "B3052_PAP3001_Teil_erkannt".
   // Fällt ab sobald das Objekt fertig zusammen gebaut ist über das Signal "Teil fertig".
   // Prüft Stop bedingung.
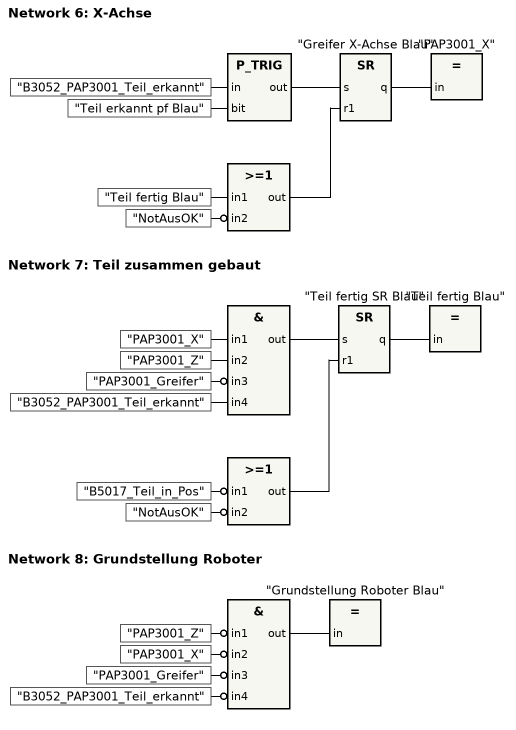
   #_w1 := "B3052_PAP3001_Teil_erkannt" AND NOT "Teil erkannt pf Blau";   // rising edge
   "Teil erkannt pf Blau" := "B3052_PAP3001_Teil_erkannt";
   IF #_w1 THEN
       "Greifer X-Achse Blau" := TRUE;   // SR flip-flop
   END_IF;
   IF "Teil fertig Blau" OR NOT "NotAusOK" THEN "Greifer X-Achse Blau" := FALSE; END_IF;
   "PAP3001_X" := "Greifer X-Achse Blau";
END_REGION

REGION Network 7: Teil zusammen gebaut
   // Der zusammen bau ist beendet wenn folgende Positionslagen erreicht sind.
   // Somit wird der Merker "Teil fertig" aktiviert und gibt das Signal für die Weitergabe an die Kommissionierung.
   // Prüft Stop bedingung.
   IF "PAP3001_X" AND "PAP3001_Z" AND NOT "PAP3001_Greifer" AND "B3052_PAP3001_Teil_erkannt" THEN
       "Teil fertig SR Blau" := TRUE;   // SR flip-flop
   END_IF;
   IF NOT "B5017_Teil_in_Pos" OR NOT "NotAusOK" THEN "Teil fertig SR Blau" := FALSE; END_IF;
   "Teil fertig Blau" := "Teil fertig SR Blau";
END_REGION

REGION Network 8: Grundstellung Roboter
   // Merker "Grundstellung Roboter" wird aktiv wenn alle Aktoren des Roboters aus sind.
   "Grundstellung Roboter Blau" := NOT "PAP3001_Z" AND NOT "PAP3001_X" AND NOT "PAP3001_Greifer" AND NOT "B3052_PAP3001_Teil_erkannt";
END_REGION
END_FUNCTION_BLOCK

FUNCTION_BLOCK "05_Weitergabe"   // FB6, FBD
{ S7_Optimized_Access := 'FALSE' }
VERSION : 0.1
BEGIN

REGION Network 1: Freigabe zur Kommissionierung
   // Der Aktor "POS3001_Heben" öffnet/schließt die Weitergabe zur Kommissionierung
   // Wird erst aktiv wenn "Teil fertig" und "Grundstellung Roboter" ein Signal liefern,
   // und setzte den Merker "FreigabeKommissionierung" (was TB3001 aktiviert ).
   // Beides fällt ab, wenn der Sensor "B3001_TB3001" unterbrochen wird.
   // Prüft Start/Stop bedingungen.
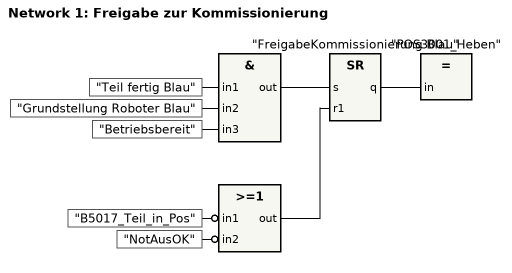
   IF "Teil fertig Blau" AND "Grundstellung Roboter Blau" AND "Betriebsbereit" THEN
       "FreigabeKommissionierung Blau" := TRUE;   // SR flip-flop
   END_IF;
   IF NOT "B5017_Teil_in_Pos" OR NOT "NotAusOK" THEN "FreigabeKommissionierung Blau" := FALSE; END_IF;
   "POS3001_Heben" := "FreigabeKommissionierung Blau";
END_REGION
END_FUNCTION_BLOCK

FUNCTION_BLOCK "06_Auswahl OT_UT"   // FB7, FBD
{ S7_Optimized_Access := 'FALSE' }
VERSION : 0.1
BEGIN

REGION Network 1: Fertigungszentrum Auswahl Unterteil/Oberteil UT =0 / OT=1
   // Signal zum erzeugen eines Oberteils.
   // Wechselndes Signal nach jeder Bearbeitung über die Sensoren "B3007_UT_BL" und "B3008_OT_BL".
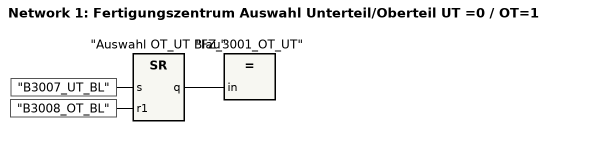
   IF "B3007_UT_BL" THEN
       "Auswahl OT_UT Blau" := TRUE;   // SR flip-flop
   END_IF;
   IF "B3008_OT_BL" THEN "Auswahl OT_UT Blau" := FALSE; END_IF;
   "FZ_3001_OT_UT" := "Auswahl OT_UT Blau";
END_REGION
END_FUNCTION_BLOCK

FUNCTION_BLOCK "02_Bearbeitung"   // FB16, FBD
{ S7_Optimized_Access := 'FALSE' }
VERSION : 0.1
   VAR
      IEC_Timer_0_Instance : TON;
      IEC_Timer_1_Instance : TOF;
   END_VAR
BEGIN

REGION Network 1: Teilbearbeiten
   // Der Merker "Signal_Start_Bearbeitung"der von Sensor "B3010_TB3007"gesteuert wird, gibt ein Signal an den Timer.
   // Nach kurzer verzögerung T#0.5s beginnt der Roboter die Bearbeitung."FZ_3001_Start"
   // Prüft Start bedingungen.
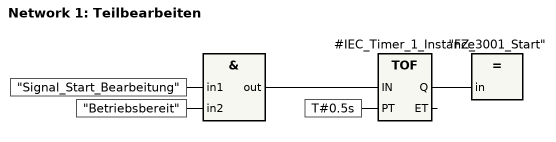
   #IEC_Timer_1_Instance.TOF(IN := "Signal_Start_Bearbeitung" AND "Betriebsbereit", PT := T#0.5s);
   "FZ_3001_Start" := #IEC_Timer_1_Instance.Q;
END_REGION
END_FUNCTION_BLOCK

// folder: Montage/Bearbeitung Grün

FUNCTION_BLOCK "01Transportband vor Bearbeitung Grün"   // FB8, FBD
{ S7_Optimized_Access := 'FALSE' }
VERSION : 0.1
   VAR_TEMP   // added for the SCL form of the ladder/FBD networks
      _w1 : Bool;
   END_VAR
BEGIN

REGION Network 1: "TB4008"
   // Prüft Start/Stop bedingungen 
   // Band 3008 Start nachdem Sensor "B3013_TB3008" unterbrochen wird.
   // Stoppt wenn Sensor "B3011_TB3007" unterbrochen wird.
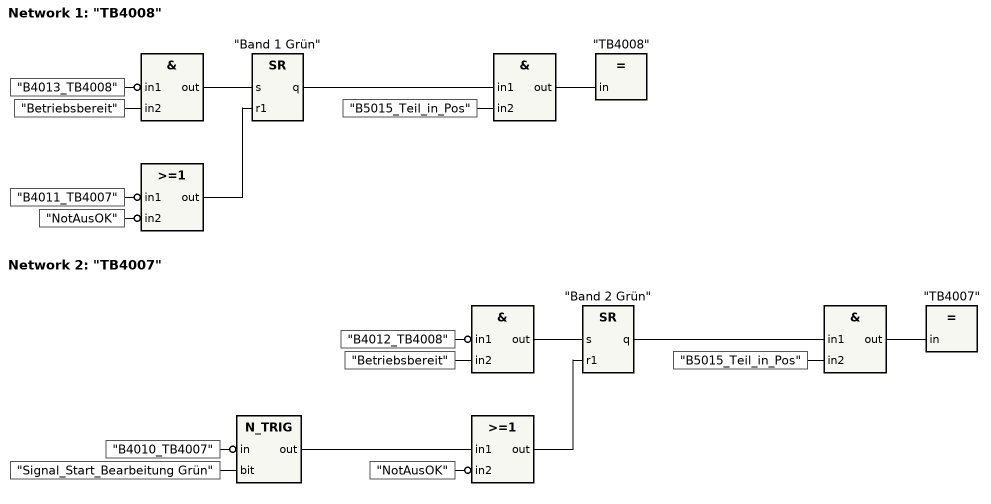
   IF NOT "B4013_TB4008" AND "Betriebsbereit" THEN
       "Band 1 Grün" := TRUE;   // SR flip-flop
   END_IF;
   IF NOT "B4011_TB4007" OR NOT "NotAusOK" THEN "Band 1 Grün" := FALSE; END_IF;
   "TB4008" := "Band 1 Grün" AND "B5015_Teil_in_Pos";
END_REGION

REGION Network 2: "TB4007"
   // Band 4007 Start nachem Sensor "B4012_TB4008" unterbrochen wird.
   // Fällt ab wenn Sensor "B4010_TB4007" unterbrochen wird.
   // Sensor "B4010_TB4007" erzeugt ein Signal für die Weiterverarbeitung:"Signal_Start_Bearbeitung Grün"
   // Prüft Start/Stop bedingungen
   #_w1 := NOT (NOT "B4010_TB4007") AND "Signal_Start_Bearbeitung Grün";   // falling edge
   "Signal_Start_Bearbeitung Grün" := NOT "B4010_TB4007";
   IF NOT "B4012_TB4008" AND "Betriebsbereit" THEN
       "Band 2 Grün" := TRUE;   // SR flip-flop
   END_IF;
   IF #_w1 OR NOT "NotAusOK" THEN "Band 2 Grün" := FALSE; END_IF;
   "TB4007" := "Band 2 Grün" AND "B5015_Teil_in_Pos";
END_REGION
END_FUNCTION_BLOCK

FUNCTION_BLOCK "02_Bearbeitung Grün"   // FB10, FBD
{ S7_Optimized_Access := 'FALSE' }
VERSION : 0.1
   VAR
      IEC_Timer_0_Instance : TON;
      IEC_Timer_1_Instance : TOF;
      IEC_Timer_2_Instance : TOF;
   END_VAR
BEGIN

REGION Network 1: Teilbearbeiten
   // Der Merker "Signal_Start_Bearbeitung"der von Sensor "B4010_TB4007"gesteuert wird, gibt ein Signal an den Timer.
   // Nach kurzer verzögerung T#0.5s beginnt der Roboter die Bearbeitung."FZ_4001_Start"
   // Prüft Start bedingungen.
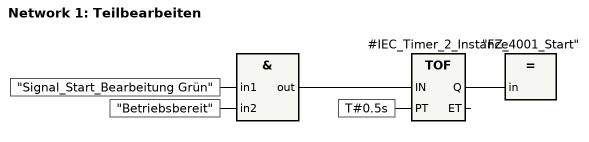
   #IEC_Timer_2_Instance.TOF(IN := "Signal_Start_Bearbeitung Grün" AND "Betriebsbereit", PT := T#0.5s);
   "FZ_4001_Start" := #IEC_Timer_2_Instance.Q;
END_REGION
END_FUNCTION_BLOCK

FUNCTION_BLOCK "03_Weiterverarbeitung Grün"   // FB11, FBD
{ S7_Optimized_Access := 'FALSE' }
VERSION : 0.1
   VAR_TEMP   // added for the SCL form of the ladder/FBD networks
      _w1 : Bool;
   END_VAR
BEGIN

REGION Network 1: "TB4006"
   // Band 4006 Start wenn Sensor "B4009_TB4006" unterbrochen wird.
   // Stoppt wenn Sensor "B4004_TB4001" oder "B4014_TB4005" unterbrochen wird.
   // Prüft Start/Stop bedingungen.
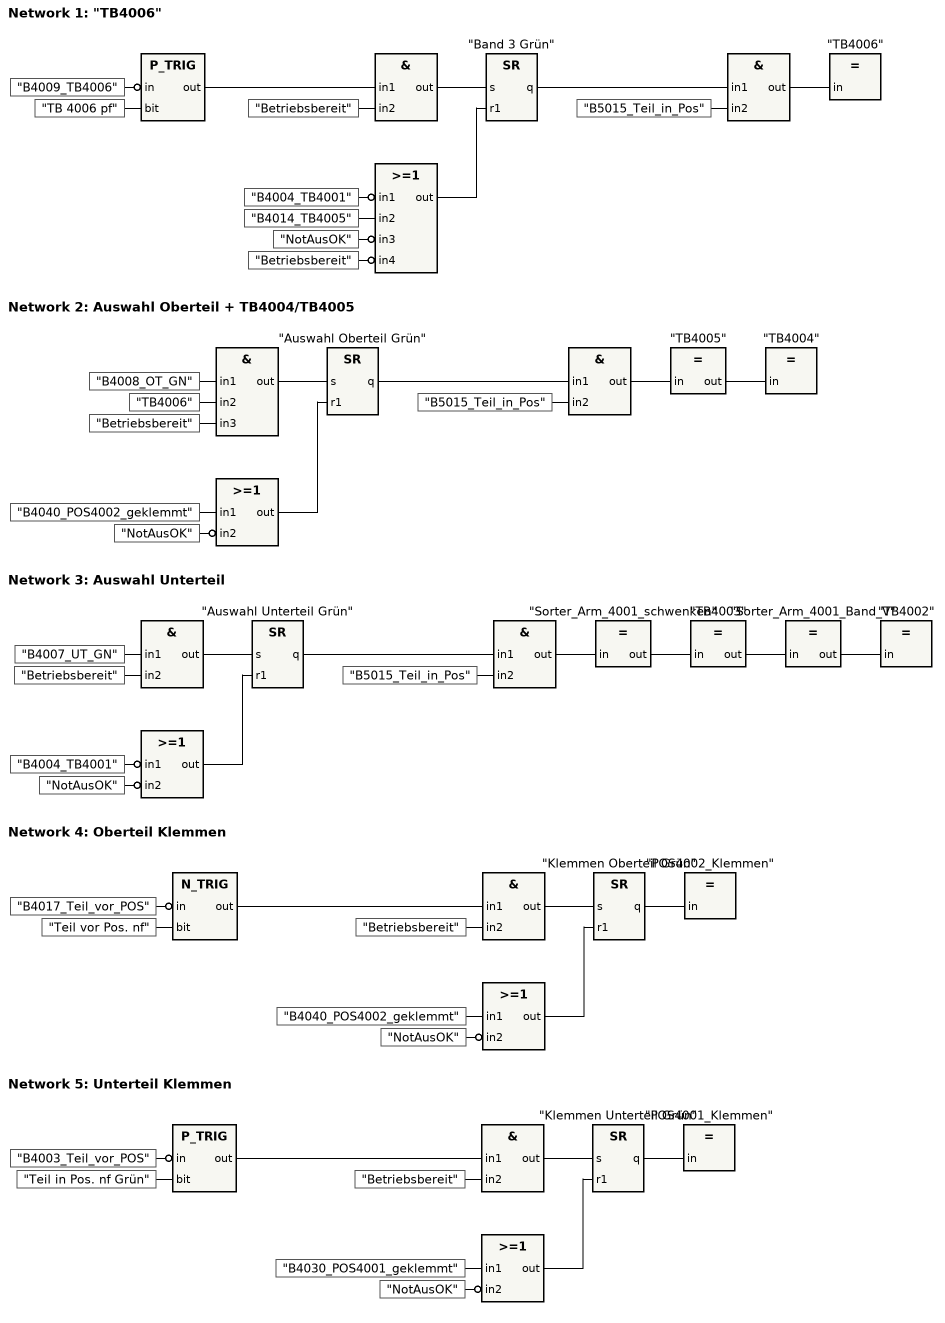
   #_w1 := NOT "B4009_TB4006" AND NOT "TB 4006 pf";   // rising edge
   "TB 4006 pf" := NOT "B4009_TB4006";
   IF #_w1 AND "Betriebsbereit" THEN
       "Band 3 Grün" := TRUE;   // SR flip-flop
   END_IF;
   IF NOT "B4004_TB4001" OR "B4014_TB4005" OR NOT "NotAusOK" OR NOT "Betriebsbereit" THEN
       "Band 3 Grün" := FALSE;
   END_IF;
   "TB4006" := "Band 3 Grün" AND "B5015_Teil_in_Pos";
END_REGION

REGION Network 2: Auswahl Oberteil + TB4004/TB4005
   // Band "TB4005" und "TB4004" starten wenn der Sensor "B4008_OT_GN" und das Band "TB4006" aktiv ist.
   // Setzt sich zurück sobald Objekt geklemmt wurde mit dem Sensor "B4040_POS4002_geklemmt".
   // Prüft Start/Stop bedingungen.
   IF "B4008_OT_GN" AND "TB4006" AND "Betriebsbereit" THEN
       "Auswahl Oberteil Grün" := TRUE;   // SR flip-flop
   END_IF;
   IF "B4040_POS4002_geklemmt" OR NOT "NotAusOK" THEN "Auswahl Oberteil Grün" := FALSE; END_IF;
   "TB4005" := "Auswahl Oberteil Grün" AND "B5015_Teil_in_Pos";
   "TB4004" := "TB4005";
END_REGION

REGION Network 3: Auswahl Unterteil
   // "Sorter_Arm_4001_schwenken","TB4003","Sorter_Arm_4001_Band_V","TB4002" werden aktiv sobald 
   // Sensor "B4007_UT_GN" reagiert.
   // Setzt sich zurück sobald das Objekt den Sensor "B4004_TB4001" unterbricht.
   // Prüft Start/Stop bedingungen.
   IF "B4007_UT_GN" AND "Betriebsbereit" THEN
       "Auswahl Unterteil Grün" := TRUE;   // SR flip-flop
   END_IF;
   IF NOT "B4004_TB4001" OR NOT "NotAusOK" THEN "Auswahl Unterteil Grün" := FALSE; END_IF;
   "Sorter_Arm_4001_schwenken" := "Auswahl Unterteil Grün" AND "B5015_Teil_in_Pos";
   "TB4003" := "Sorter_Arm_4001_schwenken";
   "Sorter_Arm_4001_Band_V" := "Sorter_Arm_4001_schwenken";
   "TB4002" := "Sorter_Arm_4001_schwenken";
END_REGION

REGION Network 4: Oberteil Klemmen
   // Objekt wird geklemmt sobald es den Sensor "B4017_Teil_vor_POS" unterbricht.
   // Fällt ab sobald Objekt geklemmt wurde: "B4040_POS4002_geklemmt".
   // Prüft Start/Stop bedingungen.
   #_w1 := NOT (NOT "B4017_Teil_vor_POS") AND "Teil vor Pos. nf";   // falling edge
   "Teil vor Pos. nf" := NOT "B4017_Teil_vor_POS";
   IF #_w1 AND "Betriebsbereit" THEN
       "Klemmen Oberteil Grün" := TRUE;   // SR flip-flop
   END_IF;
   IF "B4040_POS4002_geklemmt" OR NOT "NotAusOK" THEN "Klemmen Oberteil Grün" := FALSE; END_IF;
   "POS4002_Klemmen" := "Klemmen Oberteil Grün";
END_REGION

REGION Network 5: Unterteil Klemmen
   // Objekt wird geklemmt sobald es den Sensor "B4003_Teil_vor_POS" unterbricht.
   // Fällt ab sobald Objekt geklemmt wurde:"B4030_POS4001_geklemmt".
   // Prüft Start/Stop bedingungen.
   #_w1 := NOT "B4003_Teil_vor_POS" AND NOT "Teil in Pos. nf Grün";   // rising edge
   "Teil in Pos. nf Grün" := NOT "B4003_Teil_vor_POS";
   IF #_w1 AND "Betriebsbereit" THEN
       "Klemmen Unterteil Grün" := TRUE;   // SR flip-flop
   END_IF;
   IF "B4030_POS4001_geklemmt" OR NOT "NotAusOK" THEN "Klemmen Unterteil Grün" := FALSE; END_IF;
   "POS4001_Klemmen" := "Klemmen Unterteil Grün";
END_REGION

REGION Network 6: Unterteil TB4001 bis zur Klemme
   // Wenn Sensor "B4005_TB4002" unterbrochen wird oder das Signal "FreigabeKommissionierung" aktiviert sich "TB4001".
   // Fällt ab wenn das Objekt geklemmt wurde.
   // Prüft Start/Stop bedingungen.
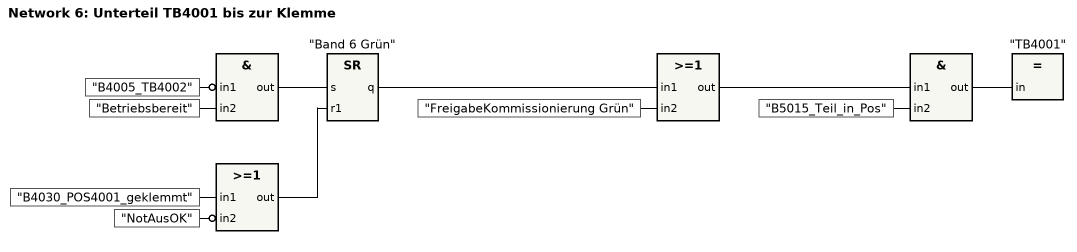
   IF NOT "B4005_TB4002" AND "Betriebsbereit" THEN
       "Band 6 Grün" := TRUE;   // SR flip-flop
   END_IF;
   IF "B4030_POS4001_geklemmt" OR NOT "NotAusOK" THEN "Band 6 Grün" := FALSE; END_IF;
   "TB4001" := ("Band 6 Grün" OR "FreigabeKommissionierung Grün") AND "B5015_Teil_in_Pos";
END_REGION
END_FUNCTION_BLOCK

FUNCTION_BLOCK "04_Zusammenbau Grün"   // FB12, FBD
{ S7_Optimized_Access := 'FALSE' }
VERSION : 0.1
   VAR_TEMP   // added for the SCL form of the ladder/FBD networks
      _w1 : Bool;
      _w2 : Bool;
      _w3 : Bool;
   END_VAR
BEGIN

REGION Network 1: Prüfung Unterteil vorhanden
   // Merker "Freigabe_Zusammenbau UT" wird gesetzt wenn das Objekt geklemmt wurde."POS4001_Klemmen"
   // Fällt ab sobald das fertige Objekt in die Kommissionierung weiter gegeben wurde."B4001_TB4001"
   // Prüft Start/Stop bedingungen.
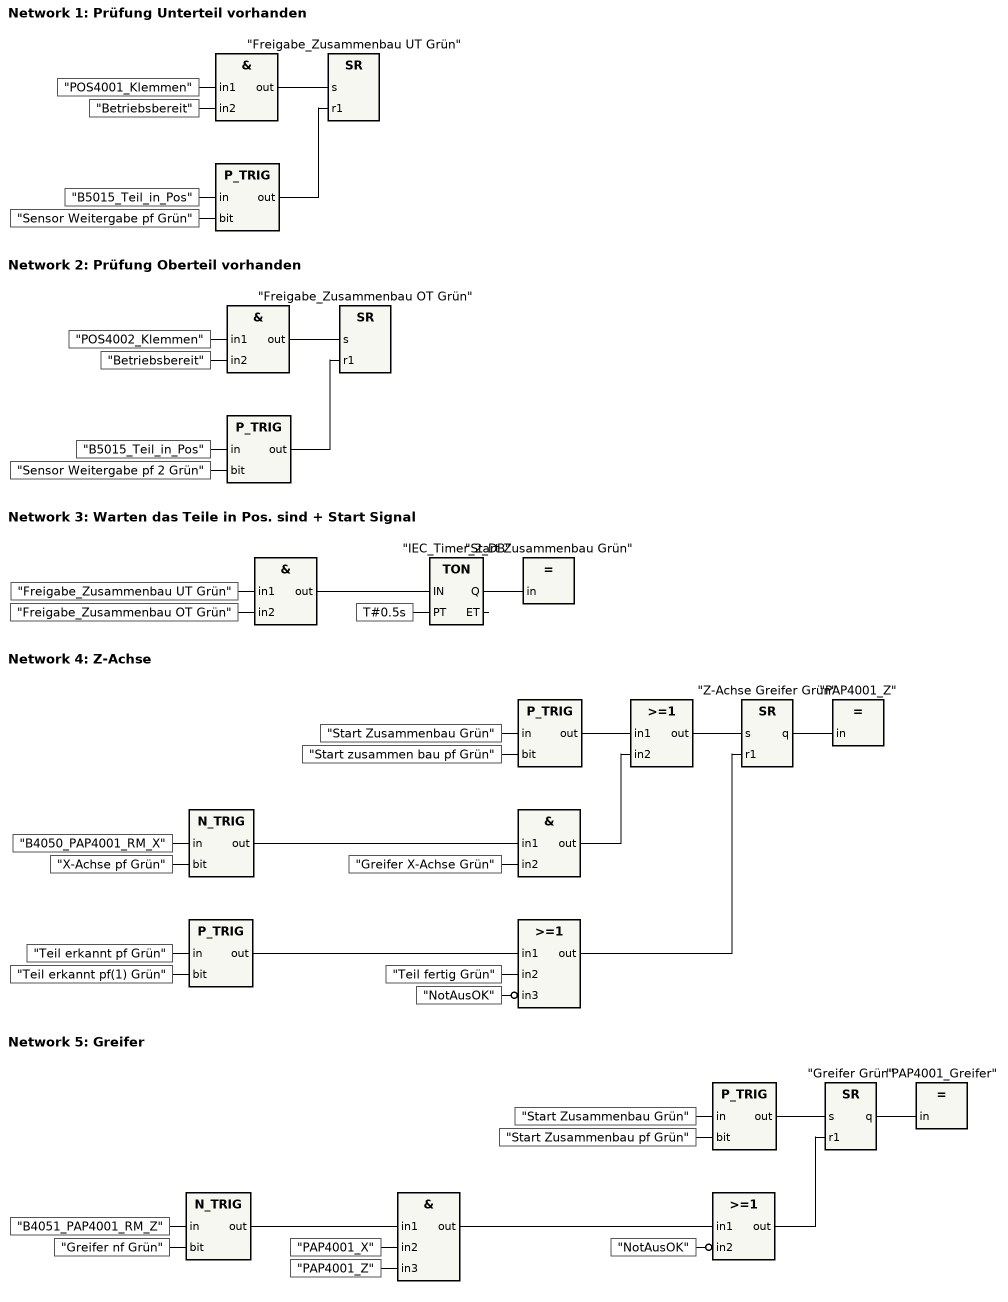
   #_w1 := "B5015_Teil_in_Pos" AND NOT "Sensor Weitergabe pf Grün";   // rising edge
   "Sensor Weitergabe pf Grün" := "B5015_Teil_in_Pos";
   IF "POS4001_Klemmen" AND "Betriebsbereit" THEN
       "Freigabe_Zusammenbau UT Grün" := TRUE;   // SR flip-flop
   END_IF;
   IF #_w1 THEN "Freigabe_Zusammenbau UT Grün" := FALSE; END_IF;
END_REGION

REGION Network 2: Prüfung Oberteil vorhanden
   // Merker"Freigabe_Zusammenbau OT" wird gesetzt wenn das Objekt geklemmt wurde."POS4002_Klemmen"
   // Fällt ab sobald das fertige Objekt in die Kommissionierung weiter gegeben wurde."B4001_TB4001"
   // Prüft Start/Stop bedingungen.
   #_w1 := "B5015_Teil_in_Pos" AND NOT "Sensor Weitergabe pf 2 Grün";   // rising edge
   "Sensor Weitergabe pf 2 Grün" := "B5015_Teil_in_Pos";
   IF "POS4002_Klemmen" AND "Betriebsbereit" THEN
       "Freigabe_Zusammenbau OT Grün" := TRUE;   // SR flip-flop
   END_IF;
   IF #_w1 THEN "Freigabe_Zusammenbau OT Grün" := FALSE; END_IF;
END_REGION

REGION Network 3: Warten das Teile in Pos. sind + Start Signal
   // Sobald beide Freigaben erteilt wurden, wird nach T#0.5s das Signal "Start Zusammenbau" erzeugt.
   "IEC_Timer_2_DB".TON(IN := "Freigabe_Zusammenbau UT Grün" AND "Freigabe_Zusammenbau OT Grün", PT := T#0.5s);
   "Start Zusammenbau Grün" := "IEC_Timer_2_DB".Q;
END_REGION

REGION Network 4: Z-Achse
   // Z-Achse senkt sich sobald das Startsignal "Start Zusammenbau" aktiv ist.
   // Fähr hoch wenn ein Teil erkannt wurde "Teil erkannt pf"oder das das Signal "Teil fertig" kommt.
   // Prüft Start/Stop bedingungen.
   #_w1 := "Start Zusammenbau Grün" AND NOT "Start zusammen bau pf Grün";   // rising edge
   "Start zusammen bau pf Grün" := "Start Zusammenbau Grün";
   #_w2 := NOT "B4050_PAP4001_RM_X" AND "X-Achse pf Grün";   // falling edge
   "X-Achse pf Grün" := "B4050_PAP4001_RM_X";
   #_w3 := "Teil erkannt pf Grün" AND NOT "Teil erkannt pf(1) Grün";   // rising edge
   "Teil erkannt pf(1) Grün" := "Teil erkannt pf Grün";
   IF #_w1 OR (#_w2 AND "Greifer X-Achse Grün") THEN
       "Z-Achse Greifer Grün" := TRUE;   // SR flip-flop
   END_IF;
   IF #_w3 OR "Teil fertig Grün" OR NOT "NotAusOK" THEN "Z-Achse Greifer Grün" := FALSE; END_IF;
   "PAP4001_Z" := "Z-Achse Greifer Grün";
END_REGION

REGION Network 5: Greifer
   // Greifer wird aktiviert sobald das Signal "Start Zusammenbau"kommt.
   // Fällt ab sobald das Objekt fertig zusammen gebaut ist über das Signal "B4051_PAP4001_RM_Z" wenn die jeweiligen X und Z Achsenposition
   // des Roboterarms entsprechend positioniert sind."PAP4001_X","PAP4001_Z".
   // Prüft Stop bedingung.
   #_w1 := "Start Zusammenbau Grün" AND NOT "Start Zusammenbau pf Grün";   // rising edge
   "Start Zusammenbau pf Grün" := "Start Zusammenbau Grün";
   #_w2 := NOT "B4051_PAP4001_RM_Z" AND "Greifer nf Grün";   // falling edge
   "Greifer nf Grün" := "B4051_PAP4001_RM_Z";
   IF #_w1 THEN
       "Greifer Grün" := TRUE;   // SR flip-flop
   END_IF;
   IF (#_w2 AND "PAP4001_X" AND "PAP4001_Z") OR NOT "NotAusOK" THEN "Greifer Grün" := FALSE; END_IF;
   "PAP4001_Greifer" := "Greifer Grün";
END_REGION

REGION Network 6: X-Achse
   // Z-Achse fährt aus sobald ein Teil erkannt wurde "B4052_PAP4001_Teil_erkannt".
   // Fällt ab sobald das Objekt fertig zusammen gebaut ist über das Signal "Teil fertig Grün".
   // Prüft Stop bedingung.
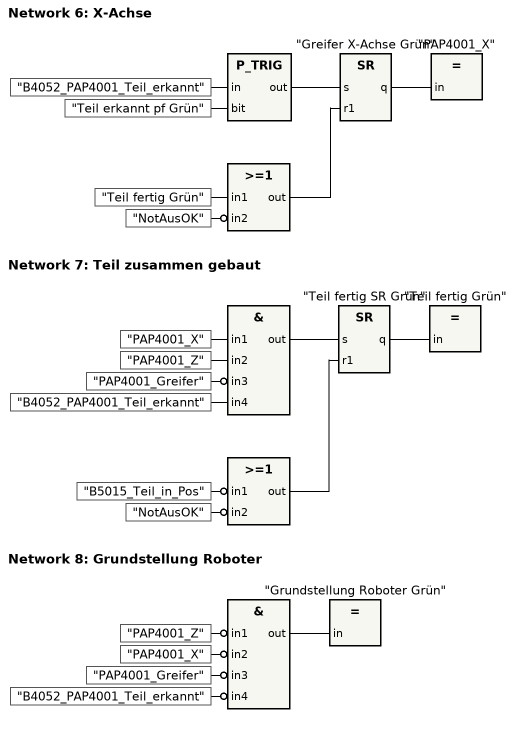
   #_w1 := "B4052_PAP4001_Teil_erkannt" AND NOT "Teil erkannt pf Grün";   // rising edge
   "Teil erkannt pf Grün" := "B4052_PAP4001_Teil_erkannt";
   IF #_w1 THEN
       "Greifer X-Achse Grün" := TRUE;   // SR flip-flop
   END_IF;
   IF "Teil fertig Grün" OR NOT "NotAusOK" THEN "Greifer X-Achse Grün" := FALSE; END_IF;
   "PAP4001_X" := "Greifer X-Achse Grün";
END_REGION

REGION Network 7: Teil zusammen gebaut
   // Der zusammen bau ist beendet wenn folgende Positionslagen erreicht sind.
   // Somit wird der Merker "Teil fertig" aktiviert und gibt das Signal für die Weitergabe an die Kommissionierung.
   // Prüft Stop bedingung.
   IF "PAP4001_X" AND "PAP4001_Z" AND NOT "PAP4001_Greifer" AND "B4052_PAP4001_Teil_erkannt" THEN
       "Teil fertig SR Grün" := TRUE;   // SR flip-flop
   END_IF;
   IF NOT "B5015_Teil_in_Pos" OR NOT "NotAusOK" THEN "Teil fertig SR Grün" := FALSE; END_IF;
   "Teil fertig Grün" := "Teil fertig SR Grün";
END_REGION

REGION Network 8: Grundstellung Roboter
   // Merker "Grundstellung Roboter" wird aktiv wenn alle Aktoren des Roboters aus sind.
   "Grundstellung Roboter Grün" := NOT "PAP4001_Z" AND NOT "PAP4001_X" AND NOT "PAP4001_Greifer" AND NOT "B4052_PAP4001_Teil_erkannt";
END_REGION
END_FUNCTION_BLOCK

FUNCTION_BLOCK "05_Weitergabe Grün"   // FB13, FBD
{ S7_Optimized_Access := 'FALSE' }
VERSION : 0.1
BEGIN

REGION Network 1: Freigabe zur Kommissionierung
   // Der Aktor "POS4001_Heben" öffnet/schließt die Weitergabe zur Kommissionierung
   // Wird erst aktiv wenn "Teil fertig" und "Grundstellung Roboter" ein Signal liefern,
   // und setzte den Merker "FreigabeKommissionierung" (was TB4001 aktiviert ).
   // Beides fällt ab, wenn der Sensor "B4001_TB4001" unterbrochen wird.
   // Prüft Start/Stop bedingungen.
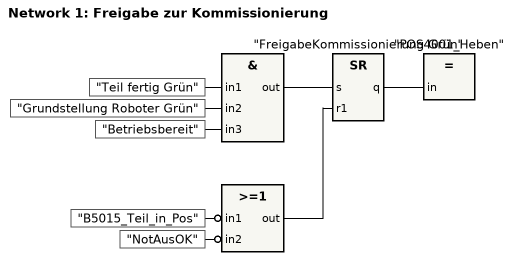
   IF "Teil fertig Grün" AND "Grundstellung Roboter Grün" AND "Betriebsbereit" THEN
       "FreigabeKommissionierung Grün" := TRUE;   // SR flip-flop
   END_IF;
   IF NOT "B5015_Teil_in_Pos" OR NOT "NotAusOK" THEN "FreigabeKommissionierung Grün" := FALSE; END_IF;
   "POS4001_Heben" := "FreigabeKommissionierung Grün";
END_REGION
END_FUNCTION_BLOCK

FUNCTION_BLOCK "06_Auswahl OT_UT_Grün"   // FB14, FBD
{ S7_Optimized_Access := 'FALSE' }
VERSION : 0.1
BEGIN

REGION Network 1: Fertigungszentrum Auswahl Unterteil/Oberteil UT =0 / OT=1
   // Signal zum erzeugen eines Oberteils.
   // Wechselndes Signal nach jeder Bearbeitung über die Sensoren "B3007_UT_BL" und "B3008_OT_BL".
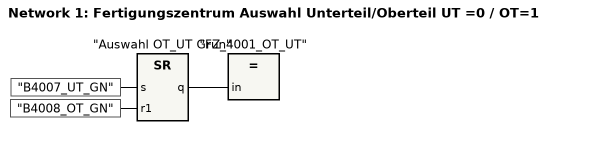
   IF "B4007_UT_GN" THEN
       "Auswahl OT_UT Grün" := TRUE;   // SR flip-flop
   END_IF;
   IF "B4008_OT_GN" THEN "Auswahl OT_UT Grün" := FALSE; END_IF;
   "FZ_4001_OT_UT" := "Auswahl OT_UT Grün";
END_REGION
END_FUNCTION_BLOCK

// folder: Montage/Bedienung

FUNCTION_BLOCK "00_Startbedingungen_2"   // FB15, FBD
{ S7_Optimized_Access := 'FALSE' }
VERSION : 0.1
   VAR_TEMP   // added for the SCL form of the ladder/FBD networks
      _w1 : Bool;
      _w2 : Bool;
   END_VAR
BEGIN

REGION Network 1: Hauptschalter
   // Anlage An + Rote Leuchte P1
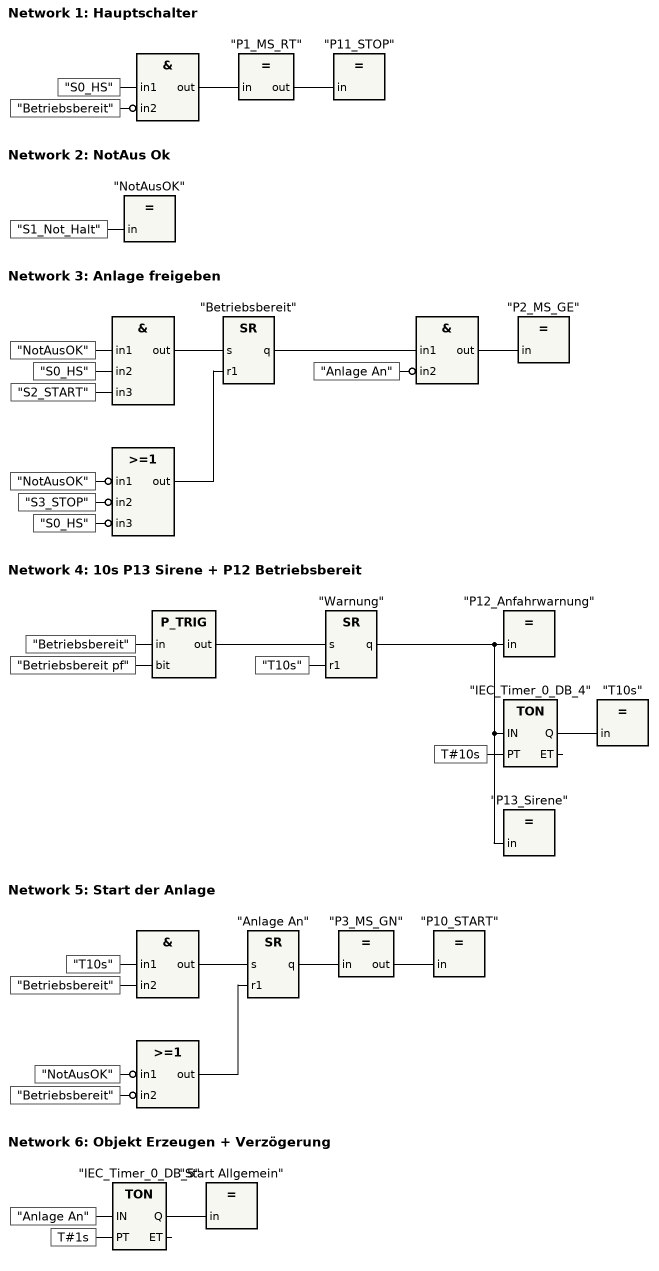
   "P1_MS_RT" := "S0_HS" AND NOT "Betriebsbereit";
   "P11_STOP" := "P1_MS_RT";
END_REGION

REGION Network 2: NotAus Ok
   // Merker NotAus Inordnung
   "NotAusOK" := "S1_Not_Halt";
END_REGION

REGION Network 3: Anlage freigeben
   // Überprüft ob Startbedingungen erfüllt sind und lässt Orange Lampe P2 zum starten leuchten.
   // "S2_START" gibt das Signal zum Starten der Anlage.
   // Freigabe der Anlage über : "Betriebsbereit"
   // Fällt ab bei: "S3_STOP","NotAusOK"
   IF "NotAusOK" AND "S0_HS" AND "S2_START" THEN
       "Betriebsbereit" := TRUE;   // SR flip-flop
   END_IF;
   IF NOT "NotAusOK" OR NOT "S3_STOP" OR NOT "S0_HS" THEN "Betriebsbereit" := FALSE; END_IF;
   "P2_MS_GE" := "Betriebsbereit" AND NOT "Anlage An";
END_REGION

REGION Network 4: 10s P13 Sirene + P12 Betriebsbereit
   // Das Signal "Betriebsbereit" setzte 10s. lang "P12_Anfahrwarnung" und "P13_Sirene" Aktiv vor dem erzeugen des ersten Objektes
   #_w1 := "Betriebsbereit" AND NOT "Betriebsbereit pf";   // rising edge
   "Betriebsbereit pf" := "Betriebsbereit";
   IF #_w1 THEN
       "Warnung" := TRUE;   // SR flip-flop
   END_IF;
   IF "T10s" THEN "Warnung" := FALSE; END_IF;
   "P12_Anfahrwarnung" := "Warnung";
   "IEC_Timer_0_DB_4".TON(IN := "Warnung", PT := T#10s);
   "T10s" := "IEC_Timer_0_DB_4".Q;
   "P13_Sirene" := "Warnung";
END_REGION

REGION Network 5: Start der Anlage
   // Sobald die Zeit abgelaufen ist wird die Grüne Leuchte Aktiv "P3_MS_GN"
   // Und der Merker "Anlage An" ist gesetzt.
   // Prüft Start/Stop bedingungen.
   IF "T10s" AND "Betriebsbereit" THEN
       "Anlage An" := TRUE;   // SR flip-flop
   END_IF;
   IF NOT "NotAusOK" OR NOT "Betriebsbereit" THEN "Anlage An" := FALSE; END_IF;
   "P3_MS_GN" := "Anlage An";
   "P10_START" := "Anlage An";
END_REGION

REGION Network 6: Objekt Erzeugen + Verzögerung
   // Nach kurzer verzögerung kommt das Startsignal: "Start Blau".
   "IEC_Timer_0_DB_5".TON(IN := "Anlage An", PT := T#1s);
   "Start Allgemein" := "IEC_Timer_0_DB_5".Q;
END_REGION

REGION Network 7: "Objekt erzeugen"
   // Da ein einfacher Flanke dem Emitter nicht reicht zum reagieren,
   // wird ein Impuls "Objekt erzeugen" von T#0.1s erzeugt.
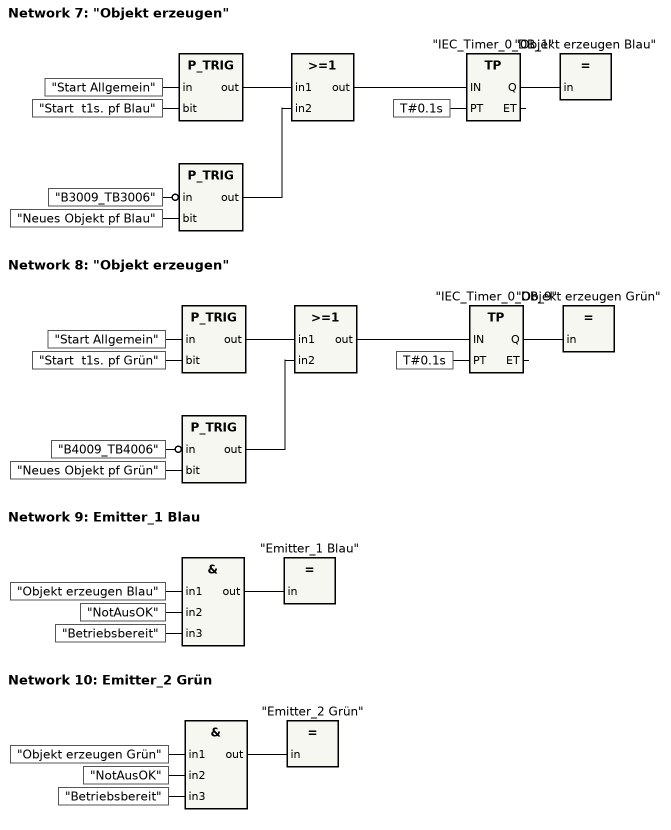
   #_w1 := "Start Allgemein" AND NOT "Start  t1s. pf Blau";   // rising edge
   "Start  t1s. pf Blau" := "Start Allgemein";
   #_w2 := NOT "B3009_TB3006" AND NOT "Neues Objekt pf Blau";   // rising edge
   "Neues Objekt pf Blau" := NOT "B3009_TB3006";
   "IEC_Timer_0_DB_1".TP(IN := #_w1 OR #_w2, PT := T#0.1s);
   "Objekt erzeugen Blau" := "IEC_Timer_0_DB_1".Q;
END_REGION

REGION Network 8: "Objekt erzeugen"
   // Da ein einfacher Flanke dem Emitter nicht reicht zum reagieren,
   // wird ein Impuls "Objekt erzeugen" von T#0.1s erzeugt.
   #_w1 := "Start Allgemein" AND NOT "Start  t1s. pf Grün";   // rising edge
   "Start  t1s. pf Grün" := "Start Allgemein";
   #_w2 := NOT "B4009_TB4006" AND NOT "Neues Objekt pf Grün";   // rising edge
   "Neues Objekt pf Grün" := NOT "B4009_TB4006";
   "IEC_Timer_0_DB_9".TP(IN := #_w1 OR #_w2, PT := T#0.1s);
   "Objekt erzeugen Grün" := "IEC_Timer_0_DB_9".Q;
END_REGION

REGION Network 9: Emitter_1 Blau
   // Prüft Start/Stop bedingungen für Emitter_1
   "Emitter_1 Blau" := "Objekt erzeugen Blau" AND "NotAusOK" AND "Betriebsbereit";
END_REGION

REGION Network 10: Emitter_2 Grün
   // Prüft Start/Stop bedingungen für Emitter_2
   "Emitter_2 Grün" := "Objekt erzeugen Grün" AND "NotAusOK" AND "Betriebsbereit";
END_REGION
END_FUNCTION_BLOCK

// ===== library: MasterCopy "RB_TB_einfach" =====

FUNCTION_BLOCK "RB_TB_einfach"   // FB101, GRAPH
{ S7_Optimized_Access := 'FALSE' }
VERSION : 0.1
// Einfacher Steuerbaustein RB / TB 
// Sensor Anfang / Ende  NO
   VAR_INPUT
      INIT_SQ : Bool := false;   // Kette in Initialzustand versetzen
      A_EIN : Bool;
      A_NOT_HALT : Bool;
      Nachfolgendes_Agg_frei : Bool;
      Sensor_vorheriges_Agg : Bool;
      Sensor_Anfang : Bool;   // Öffner
      Sensor_Ende : Bool;   // Öffner
   END_VAR
   VAR_OUTPUT
      Schritt_Nummer : Int;
      Aggregat : Bool;
      Aggregat_frei : Bool;
   END_VAR
   VAR
      HM_FLAM : Array[1..8] of Bool;
      Flanke : Array[1..8] of Bool;
      HM_Agg_Frei : Bool;
      HM_belegt : Bool;
      SWITCH : Array[0..0] of DWord;
      SW_SQTS : Array[0..6] of Byte;
      SW_ADDR : Word := 16#C;
      G7T_0 : GraphTransition;
      G7S_0 : GraphStep;
      PRE_CRIT : Array[0..1] of DWord;
      POST_CRIT : Array[0..0] of DWord;
      TVX : Array[0..2] of Byte;
      TTX : Array[0..2] of Byte;
      TSX : Array[0..2] of Byte;
      S00X : Array[0..2] of Byte;
      SOFFX : Array[0..2] of Byte;
      SONX : Array[0..2] of Byte;
      SAX : Array[0..2] of Byte;
      SERRX : Array[0..7] of Byte;
      SMX : Array[0..7] of Byte;
      S0X : Array[0..7] of Byte;
      S1X : Array[0..7] of Byte;
      S_DISPLAY : Int;   // Interne Anzeige des Ausgangsparameters S_NO
      S_SEL_OLD : Int;   // Vorheriger Wert an S_SEL
      S_DISPIDX : Byte;   // Index des Schritts, der an S_NO anliegt
      T_DISPIDX : Byte;   // Index der Transition, die an T_NO anliegt
      MOPEDGE : Struct
         AUTO : Bool := false;
         MAN : Bool := false;
         TAP : Bool := false;
         TOP : Bool := false;
         ACK_S : Bool := false;
         REG_S : Bool := false;
         T_PREV : Bool := false;
         T_NEXT : Bool := false;
         LOCK : Bool := false;
         SUP : Bool := false;
         ACKREQ : Bool := false;
         SSKIP : Bool := false;
         OFF : Bool := false;
         INIT : Bool := false;
         HALT : Bool := false;
         TMS_HALT : Bool := false;
         OPS_ZERO : Bool := false;
         SACT_DISP : Bool := false;
         SEF_DISP : Bool := false;
         SALL_DISP : Bool := false;
         S_PREV : Bool := false;
         S_NEXT : Bool := false;
         S_SELOK : Bool := false;
         S_ON : Bool := false;
         S_OFF : Bool := false;
         T_PUSH : Bool := false;
         REG : Bool := false;
         ACK : Bool := false;
         IL_PERM : Bool := false;
         T_PERM : Bool := false;
         ILP_MAN : Bool := false;
      END_STRUCT;
      MOP : Struct   // Betriebsart
         AUTO : Bool := true;   // Zustand: Automatischer Betrieb
         MAN : Bool := false;   // Zustand: Handbetrieb
         TAP : Bool := false;   // Zustand: Halbautomatisch/Weiterschalten mit Transition
         TOP : Bool := false;   // Zustand: Halbautomatisch/Ignoriere Transition
         ACK_S : Bool := false;   // Anforderung: Schritt quittieren, der an Parameter S_NO anliegt
         REG_S : Bool := false;   // Anforderung: Schritt registrieren, der an Parameter S_NO anliegt
         T_PREV : Bool := false;   // Anforderung: Vorherige gültige Transition am Parameter T_NO ausgeben
         T_NEXT : Bool := false;   // Anforderung: Nächste gültige Transition am Parameter T_NO ausgeben
         LOCK : Bool := true;   // Zustand: Interlockbearbeitung aktiviert
         SUP : Bool := true;   // Zustand: Supervisionsbearbeitung aktiviert
         ACKREQ : Bool := false;   // Zustand: Quittierung erforderlich
         SSKIP : Bool := false;   // Zustand: "Schritte überspringen" aktiviert
         OFF : Bool := false;   // Anforderung: Alle Schritte deaktivieren
         INIT : Bool := true;   // Anforderung: Kette in Initialzustand schalten
         HALT : Bool := false;   // Zustand: Kette schaltet nicht weiter
         TMS_HALT : Bool := false;   // Zustand: Alle internen Zeiten angehalten
         OPS_ZERO : Bool := false;   // Zustand: Alle mit N, L, D bearbeitete Operanden auf 0 gesetzt
         SACT_DISP : Bool := true;   // Zustand: Nur aktive Schritte anzeigen
         SEF_DISP : Bool := false;   // Zustand: Nur fehlerhafte und gestörte Schritte anzeigen
         SALL_DISP : Bool := false;   // Zustand: Alle Schritte anzeigen
         S_PREV : Bool := false;   // Anforderung: Vorherigen Schritt am Parameter S_NO ausgeben
         S_NEXT : Bool := false;   // Anforderung: Nächsten Schritt am Parameter S_NO ausgeben
         S_SELOK : Bool := false;   // Anforderung: Schrittnummer, die am Parameter S_SEL anliegt, am Parameter S_NO ausgeben
         S_ON : Bool := false;   // Anforderung: Schritt aktivieren, der am Parameter S_NO anliegt
         S_OFF : Bool := false;   // Anforderung: Schritt deaktivieren, der am Parameter S_NO anliegt
         T_PUSH : Bool := false;   // Anforderung: Schaltfreigabe für Transition
         REG : Bool := false;   // Anforderung: Alle Interlock- und Supervisionsfehler registrieren
         ACK : Bool := false;   // Anforderung: Alle Interlock- und Supervisionsfehler quittieren
         IL_PERM : Bool := false;   // Zustand: Permanente Bearbeitung aller Interlocks
         T_PERM : Bool := false;   // Zustand: Permanente Bearbeitung aller Transitionen
         ILP_MAN : Bool := false;   // Zustand: Permanente Bearbeitung aller Interlocks im Handbetrieb
      END_STRUCT;
      TICKS : Struct   // Zeittakte
         DELTA : Time := T#0ms;   // Zeitdifferenz zwischen zwei Zyklen
         OLD : Time := T#0ms;   // 10 ms Taktzählerstand im letzten Zyklus
         NEW : Time := T#0ms;   // 10 ms Taktzählerstand in diesem Zyklus
      END_STRUCT;
      SQ_FLAGS : Struct   // Kettenmerker
         ERR_FLT : Bool := false;   // Sammelfehler Interlock und Supervision
         ERROR : Bool := false;   // Sammelfehler Interlock
         FAULT : Bool := false;   // Sammelfehler Supervision
         RT_FAIL : Bool := false;   // Laufzeitfehler
         NO_SNO : Bool := false;   // Angeforderte Schrittnummer nicht gefunden
         NF_OFL : Bool := false;   // Überlauf: Zu viele Anforderungen ON oder OFF
         SA_OFL : Bool := false;   // Überlauf: Zu viele Schritte aktiv
         TV_OFL : Bool := false;   // Überlauf: Zu viele gültige Transitionen
         MSG_OFL : Bool := false;   // Überlauf: Nicht genügend Systemressourcen fü ALARM_S
         NO_SWI : Bool := false;   // Nicht Schalten in diesem Zyklus
         CYC_OP : Bool := false;   // Zyklische Bearbeitung der Kette nach Initialisierung
         AS_MSG : Bool := true;   // Meldungen zur Laufzeit durch Anweisung aktiviert oder deaktiviert
         AS_SEND : Bool := false;   // Meldungen von WR_USMSG senden oder nur in Diagnosepuffer eintragen
         SQ_BUSY : Bool := false;   // Interner Flankenmerker für Vorgangsbearbeitung
         SA_BUSY : Bool := false;   // Interner Flankenmerker für Vorgangsbearbeitung
         AS_SIG : Bool := false;   // Flankenmerker für Meldungen von Alarm_S und Alarm_SQ
      END_STRUCT;
      S_PTR : DWord := 16#450;
      S_PTR2 : DWord := 16#0;
      S_PTR3 : DWord := 16#D50;
      S_PTR4 : DWord := 16#D10;
      T_PTR : DWord := 16#CD0;
      C_AR2 : DWord := 16#0;
      M_FBDB : DWord := 16#640000;
      M_SNO : Word := 16#4;
      M_EVID : Word := 16#0;
      M_EVIL : C_Alarm_s;
      M_EVSV : C_Alarm_s;
      M_EV : DWord := 16#C30;
      CRIT : Array[0..31] of Bool;
      S_START : Byte := 16#0;
      S_IDX : Byte := 16#0;
      S_INT : Int := 72;
      S_TMP : Byte := 16#0;
      T_START : Byte := 16#0;
      T_IDX : Byte := 16#0;
      T_TMP : Byte := 16#0;
      T_TMP2 : Byte := 16#00;
      TV_POT : Byte := 16#02;
      RETURN1 : Byte := 16#0;
      RETURN2 : Byte := 16#0;
      SINI : Array[0..2] of Byte;
      LSTT : Array[0..6] of Byte;
      ATAJ : Array[0..6] of Byte;
      ATAB : Array[0..6] of Byte;
      PSTT : Array[0..6] of Byte;
      NSTT : Array[0..6] of Byte;
      ASSJ : Array[0..6] of Byte;
      ASSB : Array[0..6] of Byte;
      PTTS : Array[0..6] of Byte;
      NTTS : Array[0..6] of Byte;
      PRE_CNT : Word := 16#2;
      POST_CNT : Word := 16#1;
      ADR_COND : Word := 16#0;
      MAX_TVAL : Byte := 16#1;
      MAX_SACT : Byte := 16#1;
      MAX_CRIT : Byte := 16#4;
      T_CNT : Byte := 16#6;
      SUP_CNT : Byte := 16#0;
      LOCK_CNT : Byte := 16#5;
      S_CNT : Byte := 16#6;
      SQ_CNT : Byte := 16#1;
      PRS_INPAR : DWord := 16#40000000;
      PRS_OUTPAR : DWord := 16#0;
      GC_FLAGS : Struct
         T_MACH : Byte := 16#EB;
         COND_ED : Byte := 16#E2;
         W_LEVEL : Byte := 16#D5;
         FB_IF : Byte := 16#FA;
         AS_MSG : Word := 16#404;
         SSB : Word := 16#108;
         DILG : Word := 16#27E;
         ADDR_T0 : Word := 16#1A;
         CRIT_AVAIL : Bool := false;
         SSKIP_AVAIL : Bool := true;
         SSKIP_ON : Bool := false;
         ACK_REQ : Bool := false;
         SYNC_AVAIL : Bool := true;
         ILP_MAN : Bool := false;
         SWM_LOCKED : Bool := false;
         SAVE_SW : Bool := true;
      END_STRUCT;
      G7_FBMARK : Byte := 16#3C;
      G7_RELEASE : Byte := 16#3C;
      G7_ID2 : Byte := 16#37;
      G7_ID1 : Byte := 16#47;
   END_VAR
   // SW_SQTS[0] := 16#1;
   // TVX[0] := 16#1;
   // TTX[0] := 16#1;
   // TSX[0] := 16#1;
   // S00X[0] := 16#1;
   // SOFFX[0] := 16#1;
   // SONX[0] := 16#1;
   // SAX[0] := 16#1;
   // SERRX[0] := 16#1;
   // SMX[0] := 16#1;
   // S0X[0] := 16#1;
   // S1X[0] := 16#1;
   // SINI[0] := 16#2;
   // SINI[1] := 16#1;
   // SINI[2] := 0;
   // LSTT[0] := 0;
   // LSTT[1] := 0;
   // LSTT[2] := 0;
   // LSTT[3] := 0;
   // LSTT[4] := 0;
   // LSTT[5] := 0;
   // ATAJ[0] := 0;
   // ATAJ[1] := 16#1;
   // ATAJ[2] := 16#2;
   // ATAJ[3] := 16#3;
   // ATAJ[4] := 16#4;
   // ATAJ[5] := 16#5;
   // ATAB[0] := 0;
   // ATAB[1] := 16#1;
   // ATAB[2] := 16#2;
   // ATAB[3] := 16#3;
   // ATAB[4] := 16#4;
   // ATAB[5] := 16#5;
   // PSTT[0] := 0;
   // PSTT[1] := 16#1;
   // PSTT[2] := 16#2;
   // PSTT[3] := 16#3;
   // PSTT[4] := 16#4;
   // PSTT[5] := 16#5;
   // NSTT[0] := 16#1;
   // NSTT[1] := 16#2;
   // NSTT[2] := 16#3;
   // NSTT[3] := 16#4;
   // NSTT[4] := 16#5;
   // NSTT[5] := 16#6;
   // ASSJ[0] := 0;
   // ASSJ[1] := 16#1;
   // ASSJ[2] := 16#2;
   // ASSJ[3] := 16#3;
   // ASSJ[4] := 16#4;
   // ASSJ[5] := 16#5;
   // ASSB[0] := 0;
   // ASSB[1] := 16#1;
   // ASSB[2] := 16#2;
   // ASSB[3] := 16#3;
   // ASSB[4] := 16#4;
   // ASSB[5] := 16#5;
   // PTTS[0] := 0;
   // PTTS[2] := 16#1;
   // PTTS[3] := 16#2;
   // PTTS[4] := 16#3;
   // PTTS[5] := 16#4;
   // NTTS[0] := 0;
   // NTTS[1] := 16#1;
   // NTTS[2] := 16#2;
   // NTTS[3] := 16#3;
   // NTTS[4] := 16#4;
   // NTTS[5] := 16#5;
   // LSTT[6] := 16#1;
   // ATAJ[6] := 16#6;
   // ATAB[6] := 16#6;
   // PSTT[6] := 16#6;
   // NSTT[6] := 16#1;
   // ASSJ[6] := 16#6;
   // ASSB[6] := 16#6;
   // PTTS[6] := 16#5;
   // NTTS[6] := 16#6;
BEGIN
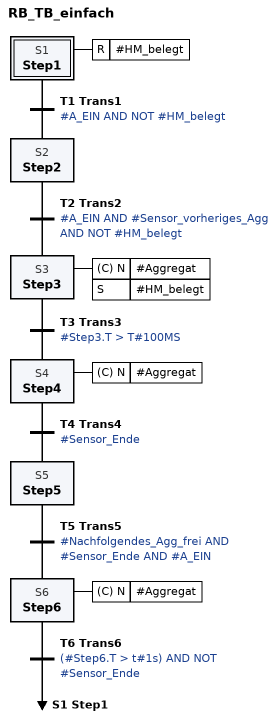
   // permanent pre-instructions
   NETWORK 1
      #HM_Agg_Frei := NOT #HM_belegt;
      #Aggregat_frei := NOT #HM_belegt;
   NETWORK 2
   TITLE = Ausgabe Schrittnummer
      #Schritt_Nummer := #S_DISPLAY;

   // sequencer 1
   INITIAL_STEP Step1:   // S1
      interlock C := NOT #A_NOT_HALT;
      // Warten auf Start
              R    #HM_belegt
   END_STEP
   TRANSITION Trans1 FROM Step1 TO Step2   // T1
      := #A_EIN AND NOT #HM_belegt;
   END_TRANSITION
   STEP Step4:   // S4
      interlock C := NOT #A_NOT_HALT;
      // Einfahrt bis Ende
      (C)     N    #Aggregat
   END_STEP
   TRANSITION Trans4 FROM Step4 TO Step5   // T4
      := #Sensor_Ende;
   END_TRANSITION
   STEP Step5:   // S5
      interlock C := NOT #A_NOT_HALT;
      // Warten auf Ausfahrt
   END_STEP
   TRANSITION Trans5 FROM Step5 TO Step6   // T5
      := #Nachfolgendes_Agg_frei AND #Sensor_Ende AND #A_EIN;
   END_TRANSITION
   STEP Step6:   // S6
      interlock C := NOT #A_NOT_HALT;
      // Ausfahrt bis Ende
      (C)     N    #Aggregat
   END_STEP
   TRANSITION Trans6 FROM Step6 TO Step1   // T6, jump
      := (#Step6.T > t#1s) AND NOT #Sensor_Ende;
   END_TRANSITION
   STEP Step3:   // S3
      interlock C := NOT #A_NOT_HALT;
      // Einfahrt Start
      (C)     N    #Aggregat
              S    #HM_belegt
   END_STEP
   TRANSITION Trans3 FROM Step3 TO Step4   // T3
      := #Step3.T > T#100MS;
   END_TRANSITION
   STEP Step2:   // S2
   END_STEP
   TRANSITION Trans2 FROM Step2 TO Step3   // T2
      := #A_EIN AND #Sensor_vorheriges_Agg AND NOT #HM_belegt;
   END_TRANSITION
END_FUNCTION_BLOCK

// ===== library: MasterCopy "Baustein_1" =====

